(* IEC 61131-3 sources: plc-st-coding-agent/progress/evidence/f14_v14_remaining_20261113/jobs/custom_minimax-m27 (part 3) *)

(* ---- public-hard-05.raw_candidate_01.st ---- *)
(* ENGINEERING_CONTRACT - Mechanical Arm Control
 * =============================================================================
 * Mode Selection: Caller ensures exactly one mode active; emergency stop has highest priority.
 *
 * Output State Table:
 * | Output          | Activation                              | Retention                     | Reset                        | Priority    |
 * |-----------------|-----------------------------------------|-------------------------------|--------------------------------|-------------|
 * | MoveDown        | Manual:DownButton AND NOT DownLimitSwitch| Manual:button hold; Auto:step | EmergencyStop, step change   | Physical dir |
 * |                 | Auto: current step = down step           | Auto: hold until limit        | button release (manual)       | rule applies |
 * | MoveUp          | Manual:UpButton AND NOT UpLimitSwitch    | Manual:button hold; Auto:step | EmergencyStop, step change   | Physical dir |
 * |                 | Auto: current step = up step             | Auto: hold until limit        | button release (manual)       | rule applies |
 * | MoveLeft        | Manual:LeftButton AND NOT LeftLimitSwitch| Manual:button hold; Auto:step | EmergencyStop, step change   | Physical dir |
 * |                 | Auto: current step = left step           | Auto: hold until limit        | button release (manual)       | rule applies |
 * | MoveRight       | Manual:RightButton AND NOT RightLimitSwitch| Manual:button hold; Auto:step| EmergencyStop, step change   | Physical dir |
 * |                 | Auto: current step = right step          | Auto: hold until limit        | button release (manual)       | rule applies |
 * | ActivateGrip    | Manual:GripButton AND NOT GripLimitSwitch| Manual:button hold; Auto:step | EmergencyStop, step change   | N/A         |
 * |                 | Auto: grip step, hold until GripLimitSwitch| Auto: hold until limit       | button release (manual)       |             |
 * | ActivateRelease | Manual:ReleaseButton AND NOT ReleaseLimitSwitch| Manual:button hold; Auto:step| EmergencyStop, step change  | N/A         |
 * |                 | Auto: release step, hold until ReleaseLimitSwitch| Auto: hold until limit    | button release (manual)       |             |
 *
 * Sequence (8 steps, single cycle and continuous modes):
 *   0: Down -> 1: Grip -> 2: Up -> 3: Right -> 4: Down -> 5: Release -> 6: Up -> 7: Left -> (repeat)
 *
 * Single step mode: Same 8-step sequence, advancing one step per Start rising edge.
 * Single cycle mode: Executes all 8 steps, stops at stepIndex=8.
 * Continuous mode: Executes all 8 steps, returns to stepIndex=0 when complete.
 *
 * Units: Limit switches TRUE=at position (normally-open, closed at position).
 * Boundary: stepIndex ∈ [0..8]; 8 = cycle complete state for single cycle mode.
 * Same-scan: Final output evaluated from current stepIndex and limit switches per scan.
 *
 * Contract PUB clauses: PUB001-PUB020 define all behavior above.
 *)

FUNCTION_BLOCK ArmController
VAR
    stepIndex : INT := 0;         // Current step in sequence (0-7), 8 = single cycle complete
    startButtonPrev : BOOL := FALSE; // Rising edge detection for Start button
    tmpRisingEdge : BOOL;
END_VAR

(* CONTRACT_RULES
[
  {"kind": "hold_until_reset", "output": "MoveDown", "set_input": "DownButton", "reset_input": null},
  {"kind": "hold_until_reset", "output": "MoveUp", "set_input": "UpButton", "reset_input": null},
  {"kind": "hold_until_reset", "output": "MoveLeft", "set_input": "LeftButton", "reset_input": null},
  {"kind": "hold_until_reset", "output": "MoveRight", "set_input": "RightButton", "reset_input": null},
  {"kind": "hold_until_reset", "output": "ActivateGrip", "set_input": "GripButton", "reset_input": null},
  {"kind": "hold_until_reset", "output": "ActivateRelease", "set_input": "ReleaseButton", "reset_input": null}
]
*)

    // Emergency stop has highest priority - stops all outputs
    IF EmergencyStop = FALSE THEN
        MoveDown := FALSE;
        MoveUp := FALSE;
        MoveLeft := FALSE;
        MoveRight := FALSE;
        ActivateGrip := FALSE;
        ActivateRelease := FALSE;
    ELSIF SingleStepMode THEN
        // Detect rising edge on Start button
        tmpRisingEdge := Start AND NOT startButtonPrev;
        startButtonPrev := Start;

        IF tmpRisingEdge THEN
            stepIndex := stepIndex + 1;
            IF stepIndex > 7 THEN
                stepIndex := 0;
            END_IF
        END_IF

        // Execute current step
        CASE stepIndex OF
            0: // Down
                MoveDown := TRUE;
                IF DownLimitSwitch THEN
                    stepIndex := 1;
                END_IF
            1: // Grip
                ActivateGrip := TRUE;
                IF GripLimitSwitch THEN
                    stepIndex := 2;
                END_IF
            2: // Up
                MoveUp := TRUE;
                IF UpLimitSwitch THEN
                    stepIndex := 3;
                END_IF
            3: // Right
                MoveRight := TRUE;
                IF RightLimitSwitch THEN
                    stepIndex := 4;
                END_IF
            4: // Down (second descent)
                MoveDown := TRUE;
                IF DownLimitSwitch THEN
                    stepIndex := 5;
                END_IF
            5: // Release
                ActivateRelease := TRUE;
                IF ReleaseLimitSwitch THEN
                    stepIndex := 6;
                END_IF
            6: // Up (second ascent)
                MoveUp := TRUE;
                IF UpLimitSwitch THEN
                    stepIndex := 7;
                END_IF
            7: // Left (return to start)
                MoveLeft := TRUE;
                IF LeftLimitSwitch THEN
                    stepIndex := 0;
                END_IF
        END_CASE

    ELSIF SingleCycleMode THEN
        // Single cycle mode: run through all steps automatically, stop at end
        CASE stepIndex OF
            0:
                MoveDown := NOT DownLimitSwitch;
                IF DownLimitSwitch THEN
                    stepIndex := 1;
                END_IF
            1:
                ActivateGrip := NOT GripLimitSwitch;
                IF GripLimitSwitch THEN
                    stepIndex := 2;
                END_IF
            2:
                MoveUp := NOT UpLimitSwitch;
                IF UpLimitSwitch THEN
                    stepIndex := 3;
                END_IF
            3:
                MoveRight := NOT RightLimitSwitch;
                IF RightLimitSwitch THEN
                    stepIndex := 4;
                END_IF
            4:
                MoveDown := NOT DownLimitSwitch;
                IF DownLimitSwitch THEN
                    stepIndex := 5;
                END_IF
            5:
                ActivateRelease := NOT ReleaseLimitSwitch;
                IF ReleaseLimitSwitch THEN
                    stepIndex := 6;
                END_IF
            6:
                MoveUp := NOT UpLimitSwitch;
                IF UpLimitSwitch THEN
                    stepIndex := 7;
                END_IF
            7:
                MoveLeft := NOT LeftLimitSwitch;
                IF LeftLimitSwitch THEN
                    stepIndex := 8; // Cycle complete, stay here
                END_IF
        END_CASE

    ELSIF ContinuousMode THEN
        // Continuous mode: run through all steps automatically, restart at end
        CASE stepIndex OF
            0:
                MoveDown := NOT DownLimitSwitch;
                IF DownLimitSwitch THEN
                    stepIndex := 1;
                END_IF
            1:
                ActivateGrip := NOT GripLimitSwitch;
                IF GripLimitSwitch THEN
                    stepIndex := 2;
                END_IF
            2:
                MoveUp := NOT UpLimitSwitch;
                IF UpLimitSwitch THEN
                    stepIndex := 3;
                END_IF
            3:
                MoveRight := NOT RightLimitSwitch;
                IF RightLimitSwitch THEN
                    stepIndex := 4;
                END_IF
            4:
                MoveDown := NOT DownLimitSwitch;
                IF DownLimitSwitch THEN
                    stepIndex := 5;
                END_IF
            5:
                ActivateRelease := NOT ReleaseLimitSwitch;
                IF ReleaseLimitSwitch THEN
                    stepIndex := 6;
                END_IF
            6:
                MoveUp := NOT UpLimitSwitch;
                IF UpLimitSwitch THEN
                    stepIndex := 7;
                END_IF
            7:
                MoveLeft := NOT LeftLimitSwitch;
                IF LeftLimitSwitch THEN
                    stepIndex := 0; // Restart cycle
                END_IF
        END_CASE

    ELSIF ManualMode THEN
        // Manual mode: direct button control with limit switch protection
        MoveDown := DownButton AND NOT DownLimitSwitch;
        MoveUp := UpButton AND NOT UpLimitSwitch;
        MoveLeft := LeftButton AND NOT LeftLimitSwitch;
        MoveRight := RightButton AND NOT RightLimitSwitch;
        ActivateGrip := GripButton AND NOT GripLimitSwitch;
        ActivateRelease := ReleaseButton AND NOT ReleaseLimitSwitch;
    END_IF

END_FUNCTION_BLOCK

(* ---- public-hard-05.raw_candidate_02.st ---- *)
(* ENGINEERING_CONTRACT - Mechanical Arm Control
 * =============================================================================
 * Mode Selection: Caller ensures exactly one mode active; emergency stop has highest priority.
 *
 * Output State Table:
 * | Output          | Activation                              | Retention                     | Reset                        | Priority    |
 * |-----------------|-----------------------------------------|-------------------------------|--------------------------------|-------------|
 * | MoveDown        | Manual:DownButton AND NOT DownLimitSwitch| Manual:button hold; Auto:step | EmergencyStop, step change   | Physical dir |
 * |                 | Auto: current step = down step           | Auto: hold until limit        | button release (manual)       | rule applies |
 * | MoveUp          | Manual:UpButton AND NOT UpLimitSwitch    | Manual:button hold; Auto:step | EmergencyStop, step change   | Physical dir |
 * |                 | Auto: current step = up step             | Auto: hold until limit        | button release (manual)       | rule applies |
 * | MoveLeft        | Manual:LeftButton AND NOT LeftLimitSwitch| Manual:button hold; Auto:step | EmergencyStop, step change   | Physical dir |
 * |                 | Auto: current step = left step           | Auto: hold until limit        | button release (manual)       | rule applies |
 * | MoveRight       | Manual:RightButton AND NOT RightLimitSwitch| Manual:button hold; Auto:step| EmergencyStop, step change   | Physical dir |
 * |                 | Auto: current step = right step          | Auto: hold until limit        | button release (manual)       | rule applies |
 * | ActivateGrip    | Manual:GripButton AND NOT GripLimitSwitch| Manual:button hold; Auto:step | EmergencyStop, step change   | N/A         |
 * |                 | Auto: grip step, hold until GripLimitSwitch| Auto: hold until limit       | button release (manual)       |             |
 * | ActivateRelease | Manual:ReleaseButton AND NOT ReleaseLimitSwitch| Manual:button hold; Auto:step| EmergencyStop, step change  | N/A         |
 * |                 | Auto: release step, hold until ReleaseLimitSwitch| Auto: hold until limit    | button release (manual)       |             |
 *
 * Sequence (8 steps, single cycle and continuous modes):
 *   0: Down -> 1: Grip -> 2: Up -> 3: Right -> 4: Down -> 5: Release -> 6: Up -> 7: Left -> (repeat)
 *
 * Single step mode: Same 8-step sequence, advancing one step per Start rising edge.
 * Single cycle mode: Executes all 8 steps, stops at stepIndex=8.
 * Continuous mode: Executes all 8 steps, returns to stepIndex=0 when complete.
 *
 * Units: Limit switches TRUE=at position (normally-open, closed at position).
 * Boundary: stepIndex ∈ [0..8]; 8 = cycle complete state for single cycle mode.
 * Same-scan: Final output evaluated from current stepIndex and limit switches per scan.
 *
 * Contract PUB clauses: PUB001-PUB020 define all behavior above.
 *)

FUNCTION_BLOCK ArmController
VAR_INPUT
    ManualMode : BOOL;
    SingleStepMode : BOOL;
    SingleCycleMode : BOOL;
    ContinuousMode : BOOL;
    EmergencyStop : BOOL;
    Start : BOOL;
    DownButton : BOOL;
    UpButton : BOOL;
    LeftButton : BOOL;
    RightButton : BOOL;
    GripButton : BOOL;
    ReleaseButton : BOOL;
    DownLimitSwitch : BOOL;
    UpLimitSwitch : BOOL;
    LeftLimitSwitch : BOOL;
    RightLimitSwitch : BOOL;
    GripLimitSwitch : BOOL;
    ReleaseLimitSwitch : BOOL;
END_VAR
VAR_OUTPUT
    MoveDown : BOOL;
    MoveUp : BOOL;
    MoveLeft : BOOL;
    MoveRight : BOOL;
    ActivateGrip : BOOL;
    ActivateRelease : BOOL;
END_VAR
VAR
    stepIndex : INT := 0;         // Current step in sequence (0-7), 8 = single cycle complete
    startButtonPrev : BOOL := FALSE; // Rising edge detection for Start button
    tmpRisingEdge : BOOL;
END_VAR

(* CONTRACT_RULES
[
  {"kind": "hold_until_reset", "output": "MoveDown", "set_input": "DownButton", "reset_input": null},
  {"kind": "hold_until_reset", "output": "MoveUp", "set_input": "UpButton", "reset_input": null},
  {"kind": "hold_until_reset", "output": "MoveLeft", "set_input": "LeftButton", "reset_input": null},
  {"kind": "hold_until_reset", "output": "MoveRight", "set_input": "RightButton", "reset_input": null},
  {"kind": "hold_until_reset", "output": "ActivateGrip", "set_input": "GripButton", "reset_input": null},
  {"kind": "hold_until_reset", "output": "ActivateRelease", "set_input": "ReleaseButton", "reset_input": null}
]
*)

    // Emergency stop has highest priority - stops all outputs
    IF EmergencyStop = FALSE THEN
        MoveDown := FALSE;
        MoveUp := FALSE;
        MoveLeft := FALSE;
        MoveRight := FALSE;
        ActivateGrip := FALSE;
        ActivateRelease := FALSE;
    ELSIF SingleStepMode THEN
        // Detect rising edge on Start button
        tmpRisingEdge := Start AND NOT startButtonPrev;
        startButtonPrev := Start;

        IF tmpRisingEdge THEN
            stepIndex := stepIndex + 1;
            IF stepIndex > 7 THEN
                stepIndex := 0;
            END_IF;
        END_IF;

        // Execute current step
        CASE stepIndex OF
            0: // Down
                MoveDown := TRUE;
                IF DownLimitSwitch THEN
                    stepIndex := 1;
                END_IF;
            1: // Grip
                ActivateGrip := TRUE;
                IF GripLimitSwitch THEN
                    stepIndex := 2;
                END_IF;
            2: // Up
                MoveUp := TRUE;
                IF UpLimitSwitch THEN
                    stepIndex := 3;
                END_IF;
            3: // Right
                MoveRight := TRUE;
                IF RightLimitSwitch THEN
                    stepIndex := 4;
                END_IF;
            4: // Down (second descent)
                MoveDown := TRUE;
                IF DownLimitSwitch THEN
                    stepIndex := 5;
                END_IF;
            5: // Release
                ActivateRelease := TRUE;
                IF ReleaseLimitSwitch THEN
                    stepIndex := 6;
                END_IF;
            6: // Up (second ascent)
                MoveUp := TRUE;
                IF UpLimitSwitch THEN
                    stepIndex := 7;
                END_IF;
            7: // Left (return to start)
                MoveLeft := TRUE;
                IF LeftLimitSwitch THEN
                    stepIndex := 0;
                END_IF;
        END_CASE;

    ELSIF SingleCycleMode THEN
        // Single cycle mode: run through all steps automatically, stop at end
        CASE stepIndex OF
            0:
                MoveDown := NOT DownLimitSwitch;
                IF DownLimitSwitch THEN
                    stepIndex := 1;
                END_IF;
            1:
                ActivateGrip := NOT GripLimitSwitch;
                IF GripLimitSwitch THEN
                    stepIndex := 2;
                END_IF;
            2:
                MoveUp := NOT UpLimitSwitch;
                IF UpLimitSwitch THEN
                    stepIndex := 3;
                END_IF;
            3:
                MoveRight := NOT RightLimitSwitch;
                IF RightLimitSwitch THEN
                    stepIndex := 4;
                END_IF;
            4:
                MoveDown := NOT DownLimitSwitch;
                IF DownLimitSwitch THEN
                    stepIndex := 5;
                END_IF;
            5:
                ActivateRelease := NOT ReleaseLimitSwitch;
                IF ReleaseLimitSwitch THEN
                    stepIndex := 6;
                END_IF;
            6:
                MoveUp := NOT UpLimitSwitch;
                IF UpLimitSwitch THEN
                    stepIndex := 7;
                END_IF;
            7:
                MoveLeft := NOT LeftLimitSwitch;
                IF LeftLimitSwitch THEN
                    stepIndex := 8; // Cycle complete, stay here
                END_IF;
        END_CASE;

    ELSIF ContinuousMode THEN
        // Continuous mode: run through all steps automatically, restart at end
        CASE stepIndex OF
            0:
                MoveDown := NOT DownLimitSwitch;
                IF DownLimitSwitch THEN
                    stepIndex := 1;
                END_IF;
            1:
                ActivateGrip := NOT GripLimitSwitch;
                IF GripLimitSwitch THEN
                    stepIndex := 2;
                END_IF;
            2:
                MoveUp := NOT UpLimitSwitch;
                IF UpLimitSwitch THEN
                    stepIndex := 3;
                END_IF;
            3:
                MoveRight := NOT RightLimitSwitch;
                IF RightLimitSwitch THEN
                    stepIndex := 4;
                END_IF;
            4:
                MoveDown := NOT DownLimitSwitch;
                IF DownLimitSwitch THEN
                    stepIndex := 5;
                END_IF;
            5:
                ActivateRelease := NOT ReleaseLimitSwitch;
                IF ReleaseLimitSwitch THEN
                    stepIndex := 6;
                END_IF;
            6:
                MoveUp := NOT UpLimitSwitch;
                IF UpLimitSwitch THEN
                    stepIndex := 7;
                END_IF;
            7:
                MoveLeft := NOT LeftLimitSwitch;
                IF LeftLimitSwitch THEN
                    stepIndex := 0; // Restart cycle
                END_IF;
        END_CASE;

    ELSIF ManualMode THEN
        // Manual mode: direct button control with limit switch protection
        MoveDown := DownButton AND NOT DownLimitSwitch;
        MoveUp := UpButton AND NOT UpLimitSwitch;
        MoveLeft := LeftButton AND NOT LeftLimitSwitch;
        MoveRight := RightButton AND NOT RightLimitSwitch;
        ActivateGrip := GripButton AND NOT GripLimitSwitch;
        ActivateRelease := ReleaseButton AND NOT ReleaseLimitSwitch;
    END_IF;

END_FUNCTION_BLOCK

(* ---- public-hard-06.candidate_01.st ---- *)
FUNCTION_BLOCK ProductionControl
VAR_INPUT
    Mode            : BOOL;
    ForwardButton   : BOOL;
    ReverseButton   : BOOL;
    SensorFeed      : BOOL;
    SensorWash      : BOOL;
    SensorWeight    : BOOL;
    SensorFiring    : BOOL;
    SensorOutput    : BOOL;
    washComplete    : BOOL;
    weightComplete  : BOOL;
    weight          : REAL;
    firingComplete  : BOOL;
END_VAR
VAR_OUTPUT
    MotorForward    : BOOL;
    MotorReverse    : BOOL;
    kick             : BOOL;
    CompletionLight : BOOL;
    firingTemp      : REAL;
END_VAR
VAR
    eState          : INT := 0;
    tmp_WashTrig    : R_TRIG;
    tmp_WeightTrig  : R_TRIG;
    tmp_FiringTrig  : R_TRIG;
    tmp_FeedPrev    : BOOL := FALSE;
END_VAR

(*
ENGINEERING_CONTRACT
================================================================================
PUB001: Mode switch (0=manual, 1=automatic)
PUB002: Manual interlocks prevent simultaneous Forward/Reverse; priority=inhibit both
PUB003: Auto sequence: FEED→WASH→WEIGH→FIRING→OUTPUT→IDLE (reset on next SensorFeed)
PUB004: Weight check [100,200]; unqualified→kick=TRUE; qualified→firingTemp=(weight-100)*0.5+500
PUB006: washComplete starts MotorForward (rising-edge, state WASH)
PUB007: weightComplete triggers weight evaluation and either kick or motor start (rising-edge)
PUB008: firingComplete starts MotorForward (rising-edge, state FIRING)
PUB010: CompletionLight := SensorOutput (retention on product presence)
PUB012: Motor stops on sensor arrival; motor starts on completion signal or qualified weight
================================================================================
Output activation table:
| Output         | Set condition                              | Reset condition        |
|----------------|--------------------------------------------|------------------------|
| MotorForward   | SensorFeed in IDLE; washComplete in WASH;  | Sensor at next station;|
|                | weightComplete in WEIGH when qualified;    | Mode change;           |
|                | firingComplete in FIRING                   | IDLE;                  |
| MotorReverse   | ReverseButton AND NOT ForwardButton; Mode=0| Mode!=0; ForwardButton |
| kick           | weightComplete in WEIGH when unqualified   | Mode change; WEIGH entry|
| CompletionLight| SensorOutput=TRUE in OUTPUT                | SensorOutput=FALSE;Mode|
| firingTemp     | weightComplete in WEIGH when qualified     | Mode change; WEIGH entry|
================================================================================
*)

tmp_FeedPrev := SensorFeed;

CASE eState OF
    0: // IDLE
        MotorForward := FALSE;
        MotorReverse := FALSE;
        kick := FALSE;
        firingTemp := 0.0;
        IF Mode = FALSE THEN
            MotorForward := ForwardButton;
            MotorReverse := (NOT ForwardButton) AND ReverseButton;
        ELSE
            IF SensorFeed AND NOT tmp_FeedPrev THEN
                MotorForward := TRUE;
                eState := 1;
            END_IF;
        END_IF;

    1: // WASH
        IF Mode = FALSE THEN
            MotorForward := FALSE;
            MotorReverse := FALSE;
            kick := FALSE;
            firingTemp := 0.0;
            eState := 0;
        ELSE
            kick := FALSE;
            firingTemp := 0.0;
            tmp_WashTrig(CLK := washComplete);
            IF SensorWash THEN
                MotorForward := FALSE;
            END_IF;
            IF tmp_WashTrig.Q THEN
                MotorForward := TRUE;
                eState := 2;
            END_IF;
        END_IF;

    2: // WEIGH
        IF Mode = FALSE THEN
            MotorForward := FALSE;
            MotorReverse := FALSE;
            kick := FALSE;
            firingTemp := 0.0;
            eState := 0;
        ELSE
            IF SensorWeight THEN
                MotorForward := FALSE;
            END_IF;
            tmp_WeightTrig(CLK := weightComplete);
            IF tmp_WeightTrig.Q THEN
                IF (weight >= 100.0) AND (weight <= 200.0) THEN
                    firingTemp := (weight - 100.0) * 0.5 + 500.0;
                    kick := FALSE;
                    MotorForward := TRUE;
                    eState := 3;
                ELSE
                    kick := TRUE;
                    firingTemp := 0.0;
                    MotorForward := TRUE;
                    eState := 3;
                END_IF;
            END_IF;
        END_IF;

    3: // FIRING
        IF Mode = FALSE THEN
            MotorForward := FALSE;
            MotorReverse := FALSE;
            kick := FALSE;
            firingTemp := 0.0;
            eState := 0;
        ELSE
            IF SensorFiring THEN
                MotorForward := FALSE;
            END_IF;
            tmp_FiringTrig(CLK := firingComplete);
            IF tmp_FiringTrig.Q THEN
                MotorForward := TRUE;
                eState := 4;
            END_IF;
        END_IF;

    4: // OUTPUT
        IF Mode = FALSE THEN
            MotorForward := FALSE;
            MotorReverse := FALSE;
            kick := FALSE;
            firingTemp := 0.0;
            CompletionLight := FALSE;
            eState := 0;
        ELSE
            IF SensorOutput THEN
                MotorForward := FALSE;
                CompletionLight := TRUE;
            ELSE
                CompletionLight := FALSE;
            END_IF;
            IF NOT SensorOutput AND (NOT MotorForward) THEN
                eState := 0;
            END_IF;
        END_IF;
END_CASE;

(* CONTRACT_RULES
[
  {"kind": "hold_until_reset", "output": "kick", "set_input": "weightComplete", "reset_input": null},
  {"kind": "hold_until_reset", "output": "firingTemp", "set_input": "weightComplete", "reset_input": null}
]
*)
END_FUNCTION_BLOCK

(* ---- public-hard-06.patch_base_02.st ---- *)
FUNCTION_BLOCK ProductionControl
VAR_INPUT
    Mode            : BOOL;
    ForwardButton   : BOOL;
    ReverseButton   : BOOL;
    SensorFeed      : BOOL;
    SensorWash      : BOOL;
    SensorWeight    : BOOL;
    SensorFiring    : BOOL;
    SensorOutput    : BOOL;
    washComplete    : BOOL;
    weightComplete  : BOOL;
    weight          : REAL;
    firingComplete  : BOOL;
END_VAR
VAR_OUTPUT
    MotorForward    : BOOL;
    MotorReverse    : BOOL;
    kick             : BOOL;
    CompletionLight : BOOL;
    firingTemp      : REAL;
END_VAR
VAR
    eState          : INT := 0;
    tmp_WashTrig    : R_TRIG;
    tmp_WeightTrig  : R_TRIG;
    tmp_FiringTrig  : R_TRIG;
    tmp_FeedPrev    : BOOL := FALSE;
END_VAR

(*
ENGINEERING_CONTRACT
================================================================================
PUB001: Mode switch (0=manual, 1=automatic)
PUB002: Manual interlocks prevent simultaneous Forward/Reverse; priority=inhibit both
PUB003: Auto sequence: FEED→WASH→WEIGH→FIRING→OUTPUT→IDLE (reset on next SensorFeed)
PUB004: Weight check [100,200]; unqualified→kick=TRUE; qualified→firingTemp=(weight-100)*0.5+500
PUB006: washComplete starts MotorForward (rising-edge, state WASH)
PUB007: weightComplete triggers weight evaluation and either kick or motor start (rising-edge)
PUB008: firingComplete starts MotorForward (rising-edge, state FIRING)
PUB010: CompletionLight := SensorOutput (retention on product presence)
PUB012: Motor stops on sensor arrival; motor starts on completion signal or qualified weight
================================================================================
Output activation table:
| Output         | Set condition                              | Reset condition        |
|----------------|--------------------------------------------|------------------------|
| MotorForward   | SensorFeed in IDLE; washComplete in WASH;  | Sensor at next station;|
|                | weightComplete in WEIGH when qualified;    | Mode change;           |
|                | firingComplete in FIRING                   | IDLE;                  |
| MotorReverse   | ReverseButton AND NOT ForwardButton; Mode=0| Mode!=0; ForwardButton |
| kick           | weightComplete in WEIGH when unqualified   | Mode change; WEIGH entry|
| CompletionLight| SensorOutput=TRUE in OUTPUT                | SensorOutput=FALSE;Mode|
| firingTemp     | weightComplete in WEIGH when qualified     | Mode change; WEIGH entry|
================================================================================
*)

tmp_FeedPrev := SensorFeed;

CASE eState OF
    0: // IDLE
        MotorForward := FALSE;
        MotorReverse := FALSE;
        kick := FALSE;
        firingTemp := 0.0;
        IF Mode = FALSE THEN
            MotorForward := ForwardButton;
            MotorReverse := (NOT ForwardButton) AND ReverseButton;
        ELSE
            IF SensorFeed AND NOT tmp_FeedPrev THEN
                MotorForward := TRUE;
                eState := 1;
            END_IF;
        END_IF;

    1: // WASH
        IF Mode = FALSE THEN
            MotorForward := FALSE;
            MotorReverse := FALSE;
            kick := FALSE;
            firingTemp := 0.0;
            eState := 0;
        ELSE
            kick := FALSE;
            firingTemp := 0.0;
            tmp_WashTrig(CLK := washComplete);
            IF SensorWash THEN
                MotorForward := FALSE;
            END_IF;
            IF tmp_WashTrig.Q THEN
                MotorForward := TRUE;
                eState := 2;
            END_IF;
        END_IF;

    2: // WEIGH
        IF Mode = FALSE THEN
            MotorForward := FALSE;
            MotorReverse := FALSE;
            kick := FALSE;
            firingTemp := 0.0;
            eState := 0;
        ELSE
            IF SensorWeight THEN
                MotorForward := FALSE;
            END_IF;
            tmp_WeightTrig(CLK := weightComplete);
            IF tmp_WeightTrig.Q THEN
                IF (weight >= 100.0) AND (weight <= 200.0) THEN
                    firingTemp := (weight - 100.0) * 0.5 + 500.0;
                    kick := FALSE;
                    MotorForward := TRUE;
                    eState := 3;
                ELSE
                    kick := TRUE;
                    firingTemp := 0.0;
                    MotorForward := TRUE;
                    eState := 3;
                END_IF;
            END_IF;
        END_IF;

    3: // FIRING
        IF Mode = FALSE THEN
            MotorForward := FALSE;
            MotorReverse := FALSE;
            kick := FALSE;
            firingTemp := 0.0;
            eState := 0;
        ELSE
            IF SensorFiring THEN
                MotorForward := FALSE;
            END_IF;
            tmp_FiringTrig(CLK := firingComplete);
            IF tmp_FiringTrig.Q THEN
                MotorForward := TRUE;
                eState := 4;
            END_IF;
        END_IF;

    4: // OUTPUT
        IF Mode = FALSE THEN
            MotorForward := FALSE;
            MotorReverse := FALSE;
            kick := FALSE;
            firingTemp := 0.0;
            CompletionLight := FALSE;
            eState := 0;
        ELSE
            IF SensorOutput THEN
                MotorForward := FALSE;
                CompletionLight := TRUE;
            ELSE
                CompletionLight := FALSE;
            END_IF;
            IF NOT SensorOutput AND (NOT MotorForward) THEN
                eState := 0;
            END_IF;
        END_IF;
END_CASE;

(* CONTRACT_RULES
[
  {"kind": "hold_until_reset", "output": "kick", "set_input": "weightComplete", "reset_input": null},
  {"kind": "hold_until_reset", "output": "firingTemp", "set_input": "weightComplete", "reset_input": null}
]
*)
END_FUNCTION_BLOCK

(* ---- public-hard-06.patch_base_03.st ---- *)
FUNCTION_BLOCK ProductionControl
VAR_INPUT
    Mode            : BOOL;
    ForwardButton   : BOOL;
    ReverseButton   : BOOL;
    SensorFeed      : BOOL;
    SensorWash      : BOOL;
    SensorWeight    : BOOL;
    SensorFiring    : BOOL;
    SensorOutput    : BOOL;
    washComplete    : BOOL;
    weightComplete  : BOOL;
    weight          : REAL;
    firingComplete  : BOOL;
END_VAR
VAR_OUTPUT
    MotorForward    : BOOL;
    MotorReverse    : BOOL;
    kick             : BOOL;
    CompletionLight : BOOL;
    firingTemp      : REAL;
END_VAR
VAR
    eState          : INT := 0;
    tmp_WashTrig    : R_TRIG;
    tmp_WeightTrig  : R_TRIG;
    tmp_FiringTrig  : R_TRIG;
    tmp_FeedPrev    : BOOL := FALSE;
END_VAR

(*
ENGINEERING_CONTRACT
================================================================================
PUB001: Mode switch (0=manual, 1=automatic)
PUB002: Manual interlocks prevent simultaneous Forward/Reverse; priority=inhibit both
PUB003: Auto sequence: FEED→WASH→WEIGH→FIRING→OUTPUT→IDLE (reset on next SensorFeed)
PUB004: Weight check [100,200]; unqualified→kick=TRUE; qualified→firingTemp=(weight-100)*0.5+500
PUB006: washComplete starts MotorForward (rising-edge, state WASH)
PUB007: weightComplete triggers weight evaluation and either kick or motor start (rising-edge)
PUB008: firingComplete starts MotorForward (rising-edge, state FIRING)
PUB010: CompletionLight := SensorOutput (retention on product presence)
PUB012: Motor stops on sensor arrival; motor starts on completion signal or qualified weight
================================================================================
Output activation table:
| Output         | Set condition                              | Reset condition        |
|----------------|--------------------------------------------|------------------------|
| MotorForward   | SensorFeed in IDLE; washComplete in WASH;  | Sensor at next station;|
|                | weightComplete in WEIGH when qualified;    | Mode change;           |
|                | firingComplete in FIRING                   | IDLE;                  |
| MotorReverse   | ReverseButton AND NOT ForwardButton; Mode=0| Mode!=0; ForwardButton |
| kick           | weightComplete in WEIGH when unqualified   | Mode change; WEIGH entry|
| CompletionLight| SensorOutput=TRUE in OUTPUT                | SensorOutput=FALSE;Mode|
| firingTemp     | weightComplete in WEIGH when qualified     | Mode change; WEIGH entry|
================================================================================
*)

tmp_FeedPrev := SensorFeed;

CASE eState OF
    0: // IDLE
        MotorForward := FALSE;
        MotorReverse := FALSE;
        kick := FALSE;
        firingTemp := 0.0;
        IF Mode = FALSE THEN
            MotorForward := ForwardButton;
            MotorReverse := (NOT ForwardButton) AND ReverseButton;
        ELSE
            IF SensorFeed AND NOT tmp_FeedPrev THEN
                MotorForward := TRUE;
                eState := 1;
            END_IF;
        END_IF;

    1: // WASH
        IF Mode = FALSE THEN
            MotorForward := FALSE;
            MotorReverse := FALSE;
            kick := FALSE;
            firingTemp := 0.0;
            eState := 0;
        ELSE
            kick := FALSE;
            firingTemp := 0.0;
            tmp_WashTrig(CLK := washComplete);
            IF SensorWash THEN
                MotorForward := FALSE;
            END_IF;
            IF tmp_WashTrig.Q THEN
                MotorForward := TRUE;
                eState := 2;
            END_IF;
        END_IF;

    2: // WEIGH
        IF Mode = FALSE THEN
            MotorForward := FALSE;
            MotorReverse := FALSE;
            kick := FALSE;
            firingTemp := 0.0;
            eState := 0;
        ELSE
            IF SensorWeight THEN
                MotorForward := FALSE;
            END_IF;
            tmp_WeightTrig(CLK := weightComplete);
            IF tmp_WeightTrig.Q THEN
                IF (weight >= 100.0) AND (weight <= 200.0) THEN
                    firingTemp := (weight - 100.0) * 0.5 + 500.0;
                    kick := FALSE;
                    MotorForward := TRUE;
                    eState := 3;
                ELSE
                    kick := TRUE;
                    firingTemp := 0.0;
                    MotorForward := TRUE;
                    eState := 3;
                END_IF;
            END_IF;
        END_IF;

    3: // FIRING
        IF Mode = FALSE THEN
            MotorForward := FALSE;
            MotorReverse := FALSE;
            kick := FALSE;
            firingTemp := 0.0;
            eState := 0;
        ELSE
            IF SensorFiring THEN
                MotorForward := FALSE;
            END_IF;
            tmp_FiringTrig(CLK := firingComplete);
            IF tmp_FiringTrig.Q THEN
                MotorForward := TRUE;
                eState := 4;
            END_IF;
        END_IF;

    4: // OUTPUT
        IF Mode = FALSE THEN
            MotorForward := FALSE;
            MotorReverse := FALSE;
            kick := FALSE;
            firingTemp := 0.0;
            CompletionLight := FALSE;
            eState := 0;
        ELSE
            IF SensorOutput THEN
                MotorForward := FALSE;
                CompletionLight := TRUE;
            ELSE
                CompletionLight := FALSE;
            END_IF;
            IF NOT SensorOutput AND (NOT MotorForward) THEN
                eState := 0;
            END_IF;
        END_IF;
END_CASE;

(* CONTRACT_RULES
[
  {"kind": "hold_until_reset", "output": "kick", "set_input": "weightComplete", "reset_input": null},
  {"kind": "hold_until_reset", "output": "firingTemp", "set_input": "weightComplete", "reset_input": null}
]
*)
END_FUNCTION_BLOCK

(* ---- public-hard-06.raw_candidate_01.st ---- *)
FUNCTION_BLOCK ProductionControl
VAR_INPUT
    Mode            : BOOL;
    ForwardButton   : BOOL;
    ReverseButton   : BOOL;
    SensorFeed      : BOOL;
    SensorWash      : BOOL;
    SensorWeight    : BOOL;
    SensorFiring    : BOOL;
    SensorOutput    : BOOL;
    washComplete    : BOOL;
    weightComplete  : BOOL;
    weight          : REAL;
    firingComplete  : BOOL;
END_VAR
VAR_OUTPUT
    MotorForward    : BOOL;
    MotorReverse    : BOOL;
    kick             : BOOL;
    CompletionLight : BOOL;
    firingTemp      : REAL;
END_VAR
VAR
    eState          : INT := 0;
    tmp_WashTrig    : R_TRIG;
    tmp_WeightTrig  : R_TRIG;
    tmp_FiringTrig  : R_TRIG;
    tmp_FeedPrev    : BOOL := FALSE;
END_VAR

(*
ENGINEERING_CONTRACT
================================================================================
PUB001: Mode switch (0=manual, 1=automatic)
PUB002: Manual interlocks prevent simultaneous Forward/Reverse; priority=inhibit both
PUB003: Auto sequence: FEED→WASH→WEIGH→FIRING→OUTPUT→IDLE (reset on next SensorFeed)
PUB004: Weight check [100,200]; unqualified→kick=TRUE; qualified→firingTemp=(weight-100)*0.5+500
PUB006: washComplete starts MotorForward (rising-edge, state WASH)
PUB007: weightComplete triggers weight evaluation and either kick or motor start (rising-edge)
PUB008: firingComplete starts MotorForward (rising-edge, state FIRING)
PUB010: CompletionLight := SensorOutput (retention on product presence)
PUB012: Motor stops on sensor arrival; motor starts on completion signal or qualified weight
================================================================================
Output activation table:
| Output         | Set condition                              | Reset condition        |
|----------------|--------------------------------------------|------------------------|
| MotorForward   | SensorFeed in IDLE; washComplete in WASH;  | Sensor at next station;|
|                | weightComplete in WEIGH when qualified;    | Mode change;           |
|                | firingComplete in FIRING                   | IDLE;                  |
| MotorReverse   | ReverseButton AND NOT ForwardButton; Mode=0| Mode!=0; ForwardButton |
| kick           | weightComplete in WEIGH when unqualified   | Mode change; WEIGH entry|
| CompletionLight| SensorOutput=TRUE in OUTPUT                | SensorOutput=FALSE;Mode|
| firingTemp     | weightComplete in WEIGH when qualified     | Mode change; WEIGH entry|
================================================================================
*)

tmp_FeedPrev := SensorFeed;

CASE eState OF
    0: // IDLE
        MotorForward := FALSE;
        MotorReverse := FALSE;
        kick := FALSE;
        firingTemp := 0.0;
        IF Mode = FALSE THEN
            MotorForward := ForwardButton;
            MotorReverse := (NOT ForwardButton) AND ReverseButton;
        ELSE
            IF SensorFeed AND NOT tmp_FeedPrev THEN
                MotorForward := TRUE;
                eState := 1;
            END_IF;
        END_IF;

    1: // WASH
        IF Mode = FALSE THEN
            MotorForward := FALSE;
            MotorReverse := FALSE;
            kick := FALSE;
            firingTemp := 0.0;
            eState := 0;
        ELSE
            kick := FALSE;
            firingTemp := 0.0;
            tmp_WashTrig(CLK := washComplete);
            IF SensorWash THEN
                MotorForward := FALSE;
            END_IF;
            IF tmp_WashTrig.Q THEN
                MotorForward := TRUE;
                eState := 2;
            END_IF;
        END_IF;

    2: // WEIGH
        IF Mode = FALSE THEN
            MotorForward := FALSE;
            MotorReverse := FALSE;
            kick := FALSE;
            firingTemp := 0.0;
            eState := 0;
        ELSE
            IF SensorWeight THEN
                MotorForward := FALSE;
            END_IF;
            tmp_WeightTrig(CLK := weightComplete);
            IF tmp_WeightTrig.Q THEN
                IF (weight >= 100.0) AND (weight <= 200.0) THEN
                    firingTemp := (weight - 100.0) * 0.5 + 500.0;
                    kick := FALSE;
                    MotorForward := TRUE;
                    eState := 3;
                ELSE
                    kick := TRUE;
                    firingTemp := 0.0;
                    MotorForward := TRUE;
                    eState := 3;
                END_IF;
            END_IF;
        END_IF;

    3: // FIRING
        IF Mode = FALSE THEN
            MotorForward := FALSE;
            MotorReverse := FALSE;
            kick := FALSE;
            firingTemp := 0.0;
            eState := 0;
        ELSE
            IF SensorFiring THEN
                MotorForward := FALSE;
            END_IF;
            tmp_FiringTrig(CLK := firingComplete);
            IF tmp_FiringTrig.Q THEN
                MotorForward := TRUE;
                eState := 4;
            END_IF;
        END_IF;

    4: // OUTPUT
        IF Mode = FALSE THEN
            MotorForward := FALSE;
            MotorReverse := FALSE;
            kick := FALSE;
            firingTemp := 0.0;
            CompletionLight := FALSE;
            eState := 0;
        ELSE
            IF SensorOutput THEN
                MotorForward := FALSE;
                CompletionLight := TRUE;
            ELSE
                CompletionLight := FALSE;
            END_IF;
            IF NOT SensorOutput AND (NOT MotorForward) THEN
                eState := 0;
            END_IF;
        END_IF;
END_CASE;

(* CONTRACT_RULES
[
  {"kind": "hold_until_reset", "output": "kick", "set_input": "weightComplete", "reset_input": null},
  {"kind": "hold_until_reset", "output": "firingTemp", "set_input": "weightComplete", "reset_input": null}
]
*)
END_FUNCTION_BLOCK

(* ---- public-medium-01.candidate_01.st ---- *)
FUNCTION_BLOCK FB_PumpControl
VAR_INPUT
    mode  : BOOL;  // FALSE: Manual, TRUE: Automatic
    start : BOOL;
    stop  : BOOL;
END_VAR

VAR_IN_OUT
    pumpGroup : ARRAY[1..5] OF ST_Pump;
END_VAR

VAR
    tmp_i          : INT;
    tmp_j          : INT;
    tmp_temp       : ST_Pump;
    tmp_tempIndex  : INT;
    tmp_sorted     : ARRAY[1..5] OF ST_Pump;
    tmp_order      : ARRAY[1..5] OF INT;
END_VAR

// ENGINEERING_CONTRACT
// ┌─────────────────────────────────────────────────────────────────────────────────────────────┐
// │ Output/State              │ Activation                   │ Retention    │ Reset/Deactivation │ Same-scan │ Boundaries      │ PUB Clause     │
// │------------------------───│──────────────────────────────│──────────────│────────────────────│───────────│─────────────────│────────────────│
// │ pumpGroup[].RunComd FALSE │ stop=TRUE                    │ -            │ start=TRUE         │ -         │ 0–5 pumps       │ PUB001, PUB004 │
// │ pumpGroup[].RunComd TRUE  │ start=TRUE AND selected only │ Hold(start)  │ stop=TRUE          │ -         │ Manual: 1–5 pumps; Auto: 3 │ PUB001, PUB003 │
// │ pumpGroup[].RunComd TRUE  │ start=TRUE AND top-3 priority│ Hold(start)  │ stop=TRUE          │ -         │ Auto: exactly 3 │ PUB002         │
// └─────────────────────────────────────────────────────────────────────────────────────────────┘

// Stop has highest priority — de-energizes all pumps immediately
IF stop THEN
    FOR tmp_i := 1 TO 5 DO
        pumpGroup[tmp_i].RunComd := FALSE;
    END_FOR;
    RETURN;
END_IF;

IF NOT mode THEN
    // Manual mode: selected pump(s) follow start command
    FOR tmp_i := 1 TO 5 DO
        IF pumpGroup[tmp_i].selection THEN
            pumpGroup[tmp_i].RunComd := start;
        ELSE
            pumpGroup[tmp_i].RunComd := FALSE;
        END_IF;
    END_FOR;
ELSE
    // Automatic mode: top-3 priority pumps follow start command
    // Copy for sorting (preserves original pumpGroup indices)
    FOR tmp_i := 1 TO 5 DO
        tmp_sorted[tmp_i] := pumpGroup[tmp_i];
        tmp_order[tmp_i]  := tmp_i;
    END_FOR;

    // Bubble sort by priority descending (stable: equal priority keeps original order)
    FOR tmp_i := 1 TO 4 DO
        FOR tmp_j := tmp_i + 1 TO 5 DO
            IF tmp_sorted[tmp_j].priority > tmp_sorted[tmp_i].priority THEN
                tmp_temp           := tmp_sorted[tmp_i];
                tmp_sorted[tmp_i]  := tmp_sorted[tmp_j];
                tmp_sorted[tmp_j]  := tmp_temp;

                tmp_tempIndex      := tmp_order[tmp_i];
                tmp_order[tmp_i]   := tmp_order[tmp_j];
                tmp_order[tmp_j]   := tmp_tempIndex;
            END_IF;
        END_FOR;
    END_FOR;

    // Enable top-3 pumps (by original index) when start is asserted
    FOR tmp_i := 1 TO 5 DO
        IF tmp_i <= 3 THEN
            pumpGroup[tmp_order[tmp_i]].RunComd := start;
        ELSE
            pumpGroup[tmp_order[tmp_i]].RunComd := FALSE;
        END_IF;
    END_FOR;
END_IF;

END_FUNCTION_BLOCK

(* CONTRACT_RULES [] *)

(* ---- public-medium-01.candidate_02.st ---- *)
TYPE ST_Pump : STRUCT
    priority  : INT;
    selection : BOOL;
    RunComd   : BOOL;
END_STRUCT
END_TYPE;

FUNCTION_BLOCK FB_PumpControl
VAR_INPUT
    mode  : BOOL;  // FALSE: Manual, TRUE: Automatic
    start : BOOL;
    stop  : BOOL;
END_VAR

VAR_IN_OUT
    pumpGroup : ARRAY[1..5] OF ST_Pump;
END_VAR

VAR
    tmp_i          : INT;
    tmp_j          : INT;
    tmp_temp       : ST_Pump;
    tmp_tempIndex  : INT;
    tmp_sorted     : ARRAY[1..5] OF ST_Pump;
    tmp_order      : ARRAY[1..5] OF INT;
END_VAR

// ENGINEERING_CONTRACT
// ┌─────────────────────────────────────────────────────────────────────────────────────────────┐
// │ Output/State              │ Activation                   │ Retention    │ Reset/Deactivation │ Same-scan │ Boundaries      │ PUB Clause     │
// │------------------------───│──────────────────────────────│──────────────│────────────────────│───────────│─────────────────│────────────────│
// │ pumpGroup[].RunComd FALSE │ stop=TRUE                    │ -            │ start=TRUE         │ -         │ 0–5 pumps       │ PUB001, PUB004 │
// │ pumpGroup[].RunComd TRUE  │ start=TRUE AND selected only │ Hold(start)  │ stop=TRUE          │ -         │ Manual: 1–5 pumps; Auto: 3 │ PUB001, PUB003 │
// │ pumpGroup[].RunComd TRUE  │ start=TRUE AND top-3 priority│ Hold(start)  │ stop=TRUE          │ -         │ Auto: exactly 3 │ PUB002         │
// └─────────────────────────────────────────────────────────────────────────────────────────────┘

// Stop has highest priority — de-energizes all pumps immediately
IF stop THEN
    FOR tmp_i := 1 TO 5 DO
        pumpGroup[tmp_i].RunComd := FALSE;
    END_FOR;
    RETURN;
END_IF;

IF NOT mode THEN
    // Manual mode: selected pump(s) follow start command
    FOR tmp_i := 1 TO 5 DO
        IF pumpGroup[tmp_i].selection THEN
            pumpGroup[tmp_i].RunComd := start;
        ELSE
            pumpGroup[tmp_i].RunComd := FALSE;
        END_IF;
    END_FOR;
ELSE
    // Automatic mode: top-3 priority pumps follow start command
    // Copy for sorting (preserves original pumpGroup indices)
    FOR tmp_i := 1 TO 5 DO
        tmp_sorted[tmp_i] := pumpGroup[tmp_i];
        tmp_order[tmp_i]  := tmp_i;
    END_FOR;

    // Bubble sort by priority descending (stable: equal priority keeps original order)
    FOR tmp_i := 1 TO 4 DO
        FOR tmp_j := tmp_i + 1 TO 5 DO
            IF tmp_sorted[tmp_j].priority > tmp_sorted[tmp_i].priority THEN
                tmp_temp           := tmp_sorted[tmp_i];
                tmp_sorted[tmp_i]  := tmp_sorted[tmp_j];
                tmp_sorted[tmp_j]  := tmp_temp;

                tmp_tempIndex      := tmp_order[tmp_i];
                tmp_order[tmp_i]   := tmp_order[tmp_j];
                tmp_order[tmp_j]   := tmp_tempIndex;
            END_IF;
        END_FOR;
    END_FOR;

    // Enable top-3 pumps (by original index) when start is asserted
    FOR tmp_i := 1 TO 5 DO
        IF tmp_i <= 3 THEN
            pumpGroup[tmp_order[tmp_i]].RunComd := start;
        ELSE
            pumpGroup[tmp_order[tmp_i]].RunComd := FALSE;
        END_IF;
    END_FOR;
END_IF;

END_FUNCTION_BLOCK

(* CONTRACT_RULES [] *)

(* ---- public-medium-01.patch_base_02.st ---- *)
FUNCTION_BLOCK FB_PumpControl
VAR_INPUT
    mode  : BOOL;  // FALSE: Manual, TRUE: Automatic
    start : BOOL;
    stop  : BOOL;
END_VAR

VAR_IN_OUT
    pumpGroup : ARRAY[1..5] OF ST_Pump;
END_VAR

VAR
    tmp_i          : INT;
    tmp_j          : INT;
    tmp_temp       : ST_Pump;
    tmp_tempIndex  : INT;
    tmp_sorted     : ARRAY[1..5] OF ST_Pump;
    tmp_order      : ARRAY[1..5] OF INT;
END_VAR

// ENGINEERING_CONTRACT
// ┌─────────────────────────────────────────────────────────────────────────────────────────────┐
// │ Output/State              │ Activation                   │ Retention    │ Reset/Deactivation │ Same-scan │ Boundaries      │ PUB Clause     │
// │------------------------───│──────────────────────────────│──────────────│────────────────────│───────────│─────────────────│────────────────│
// │ pumpGroup[].RunComd FALSE │ stop=TRUE                    │ -            │ start=TRUE         │ -         │ 0–5 pumps       │ PUB001, PUB004 │
// │ pumpGroup[].RunComd TRUE  │ start=TRUE AND selected only │ Hold(start)  │ stop=TRUE          │ -         │ Manual: 1–5 pumps; Auto: 3 │ PUB001, PUB003 │
// │ pumpGroup[].RunComd TRUE  │ start=TRUE AND top-3 priority│ Hold(start)  │ stop=TRUE          │ -         │ Auto: exactly 3 │ PUB002         │
// └─────────────────────────────────────────────────────────────────────────────────────────────┘

// Stop has highest priority — de-energizes all pumps immediately
IF stop THEN
    FOR tmp_i := 1 TO 5 DO
        pumpGroup[tmp_i].RunComd := FALSE;
    END_FOR;
    RETURN;
END_IF;

IF NOT mode THEN
    // Manual mode: selected pump(s) follow start command
    FOR tmp_i := 1 TO 5 DO
        IF pumpGroup[tmp_i].selection THEN
            pumpGroup[tmp_i].RunComd := start;
        ELSE
            pumpGroup[tmp_i].RunComd := FALSE;
        END_IF;
    END_FOR;
ELSE
    // Automatic mode: top-3 priority pumps follow start command
    // Copy for sorting (preserves original pumpGroup indices)
    FOR tmp_i := 1 TO 5 DO
        tmp_sorted[tmp_i] := pumpGroup[tmp_i];
        tmp_order[tmp_i]  := tmp_i;
    END_FOR;

    // Bubble sort by priority descending (stable: equal priority keeps original order)
    FOR tmp_i := 1 TO 4 DO
        FOR tmp_j := tmp_i + 1 TO 5 DO
            IF tmp_sorted[tmp_j].priority > tmp_sorted[tmp_i].priority THEN
                tmp_temp           := tmp_sorted[tmp_i];
                tmp_sorted[tmp_i]  := tmp_sorted[tmp_j];
                tmp_sorted[tmp_j]  := tmp_temp;

                tmp_tempIndex      := tmp_order[tmp_i];
                tmp_order[tmp_i]   := tmp_order[tmp_j];
                tmp_order[tmp_j]   := tmp_tempIndex;
            END_IF;
        END_FOR;
    END_FOR;

    // Enable top-3 pumps (by original index) when start is asserted
    FOR tmp_i := 1 TO 5 DO
        IF tmp_i <= 3 THEN
            pumpGroup[tmp_order[tmp_i]].RunComd := start;
        ELSE
            pumpGroup[tmp_order[tmp_i]].RunComd := FALSE;
        END_IF;
    END_FOR;
END_IF;

END_FUNCTION_BLOCK

(* CONTRACT_RULES [] *)

(* ---- public-medium-01.raw_candidate_01.st ---- *)
FUNCTION_BLOCK FB_PumpControl
VAR_INPUT
    mode  : BOOL;  // FALSE: Manual, TRUE: Automatic
    start : BOOL;
    stop  : BOOL;
END_VAR

VAR_IN_OUT
    pumpGroup : ARRAY[1..5] OF ST_Pump;
END_VAR

VAR
    tmp_i          : INT;
    tmp_j          : INT;
    tmp_temp       : ST_Pump;
    tmp_tempIndex  : INT;
    tmp_sorted     : ARRAY[1..5] OF ST_Pump;
    tmp_order      : ARRAY[1..5] OF INT;
END_VAR

// ENGINEERING_CONTRACT
// ┌─────────────────────────────────────────────────────────────────────────────────────────────┐
// │ Output/State              │ Activation                   │ Retention    │ Reset/Deactivation │ Same-scan │ Boundaries      │ PUB Clause     │
// │------------------------───│──────────────────────────────│──────────────│────────────────────│───────────│─────────────────│────────────────│
// │ pumpGroup[].RunComd FALSE │ stop=TRUE                    │ -            │ start=TRUE         │ -         │ 0–5 pumps       │ PUB001, PUB004 │
// │ pumpGroup[].RunComd TRUE  │ start=TRUE AND selected only │ Hold(start)  │ stop=TRUE          │ -         │ Manual: 1–5 pumps; Auto: 3 │ PUB001, PUB003 │
// │ pumpGroup[].RunComd TRUE  │ start=TRUE AND top-3 priority│ Hold(start)  │ stop=TRUE          │ -         │ Auto: exactly 3 │ PUB002         │
// └─────────────────────────────────────────────────────────────────────────────────────────────┘

// Stop has highest priority — de-energizes all pumps immediately
IF stop THEN
    FOR tmp_i := 1 TO 5 DO
        pumpGroup[tmp_i].RunComd := FALSE;
    END_FOR
    RETURN;
END_IF

IF NOT mode THEN
    // Manual mode: selected pump(s) follow start command
    FOR tmp_i := 1 TO 5 DO
        IF pumpGroup[tmp_i].selection THEN
            pumpGroup[tmp_i].RunComd := start;
        ELSE
            pumpGroup[tmp_i].RunComd := FALSE;
        END_IF
    END_FOR
ELSE
    // Automatic mode: top-3 priority pumps follow start command
    // Copy for sorting (preserves original pumpGroup indices)
    FOR tmp_i := 1 TO 5 DO
        tmp_sorted[tmp_i] := pumpGroup[tmp_i];
        tmp_order[tmp_i]  := tmp_i;
    END_FOR

    // Bubble sort by priority descending (stable: equal priority keeps original order)
    FOR tmp_i := 1 TO 4 DO
        FOR tmp_j := tmp_i + 1 TO 5 DO
            IF tmp_sorted[tmp_j].priority > tmp_sorted[tmp_i].priority THEN
                tmp_temp           := tmp_sorted[tmp_i];
                tmp_sorted[tmp_i]  := tmp_sorted[tmp_j];
                tmp_sorted[tmp_j]  := tmp_temp;

                tmp_tempIndex      := tmp_order[tmp_i];
                tmp_order[tmp_i]   := tmp_order[tmp_j];
                tmp_order[tmp_j]   := tmp_tempIndex;
            END_IF
        END_FOR
    END_FOR

    // Enable top-3 pumps (by original index) when start is asserted
    FOR tmp_i := 1 TO 5 DO
        IF tmp_i <= 3 THEN
            pumpGroup[tmp_order[tmp_i]].RunComd := start;
        ELSE
            pumpGroup[tmp_order[tmp_i]].RunComd := FALSE;
        END_IF
    END_FOR
END_IF

END_FUNCTION_BLOCK

(* CONTRACT_RULES [] *)

(* ---- public-medium-01.raw_candidate_02.st ---- *)
TYPE ST_Pump : STRUCT
    priority  : INT;
    selection : BOOL;
    RunComd   : BOOL;
END_STRUCT
END_TYPE

FUNCTION_BLOCK FB_PumpControl
VAR_INPUT
    mode  : BOOL;  // FALSE: Manual, TRUE: Automatic
    start : BOOL;
    stop  : BOOL;
END_VAR

VAR_IN_OUT
    pumpGroup : ARRAY[1..5] OF ST_Pump;
END_VAR

VAR
    tmp_i          : INT;
    tmp_j          : INT;
    tmp_temp       : ST_Pump;
    tmp_tempIndex  : INT;
    tmp_sorted     : ARRAY[1..5] OF ST_Pump;
    tmp_order      : ARRAY[1..5] OF INT;
END_VAR

// ENGINEERING_CONTRACT
// ┌─────────────────────────────────────────────────────────────────────────────────────────────┐
// │ Output/State              │ Activation                   │ Retention    │ Reset/Deactivation │ Same-scan │ Boundaries      │ PUB Clause     │
// │------------------------───│──────────────────────────────│──────────────│────────────────────│───────────│─────────────────│────────────────│
// │ pumpGroup[].RunComd FALSE │ stop=TRUE                    │ -            │ start=TRUE         │ -         │ 0–5 pumps       │ PUB001, PUB004 │
// │ pumpGroup[].RunComd TRUE  │ start=TRUE AND selected only │ Hold(start)  │ stop=TRUE          │ -         │ Manual: 1–5 pumps; Auto: 3 │ PUB001, PUB003 │
// │ pumpGroup[].RunComd TRUE  │ start=TRUE AND top-3 priority│ Hold(start)  │ stop=TRUE          │ -         │ Auto: exactly 3 │ PUB002         │
// └─────────────────────────────────────────────────────────────────────────────────────────────┘

// Stop has highest priority — de-energizes all pumps immediately
IF stop THEN
    FOR tmp_i := 1 TO 5 DO
        pumpGroup[tmp_i].RunComd := FALSE;
    END_FOR;
    RETURN;
END_IF;

IF NOT mode THEN
    // Manual mode: selected pump(s) follow start command
    FOR tmp_i := 1 TO 5 DO
        IF pumpGroup[tmp_i].selection THEN
            pumpGroup[tmp_i].RunComd := start;
        ELSE
            pumpGroup[tmp_i].RunComd := FALSE;
        END_IF;
    END_FOR;
ELSE
    // Automatic mode: top-3 priority pumps follow start command
    // Copy for sorting (preserves original pumpGroup indices)
    FOR tmp_i := 1 TO 5 DO
        tmp_sorted[tmp_i] := pumpGroup[tmp_i];
        tmp_order[tmp_i]  := tmp_i;
    END_FOR;

    // Bubble sort by priority descending (stable: equal priority keeps original order)
    FOR tmp_i := 1 TO 4 DO
        FOR tmp_j := tmp_i + 1 TO 5 DO
            IF tmp_sorted[tmp_j].priority > tmp_sorted[tmp_i].priority THEN
                tmp_temp           := tmp_sorted[tmp_i];
                tmp_sorted[tmp_i]  := tmp_sorted[tmp_j];
                tmp_sorted[tmp_j]  := tmp_temp;

                tmp_tempIndex      := tmp_order[tmp_i];
                tmp_order[tmp_i]   := tmp_order[tmp_j];
                tmp_order[tmp_j]   := tmp_tempIndex;
            END_IF;
        END_FOR;
    END_FOR;

    // Enable top-3 pumps (by original index) when start is asserted
    FOR tmp_i := 1 TO 5 DO
        IF tmp_i <= 3 THEN
            pumpGroup[tmp_order[tmp_i]].RunComd := start;
        ELSE
            pumpGroup[tmp_order[tmp_i]].RunComd := FALSE;
        END_IF;
    END_FOR;
END_IF;

END_FUNCTION_BLOCK

(* CONTRACT_RULES [] *)

(* ---- public-medium-02.candidate_01.st ---- *)
FUNCTION_BLOCK FB_AnalogBatchProcessing
VAR_INPUT
END_VAR
VAR_IN_OUT
    analogValues : ARRAY[*] OF INT;
    channels     : ARRAY[*] OF ST_AnalogChannel;
END_VAR
VAR_OUTPUT
END_VAR
VAR
END_VAR

(*
ENGINEERING_CONTRACT
================================================================================
PUB001: Process 'count' channels starting at each array's lower bound.
        Arrays passed by reference preserve caller-defined bounds.
        Read-only: analogValues elements are never modified.
PUB002: Per-channel conversion based on measuringMode field.
        - Mode 0: Linear scaling using hiLIM/loLIM and bipolar flag.
        - Mode 1: Standard temperature (raw / 10.0).
        - Mode 2: Climatic temperature (raw / 100.0).
        - Invalid mode: retVal=16#8001, outputValue unchanged.
PUB003: Mode 0 linear scaling maps raw 0..27648 (unipolar) or -27648..27648 (bipolar)
        to loLIM..hiLIM range. OutputValue = loLIM + (raw - rawMin) * (hiLIM - loLIM) / range.
PUB004: If hiLIM <= loLIM in mode 0, set retVal=16#8002 and skip conversion.
PUB005: Disabled channels (enable=FALSE) are skipped; retVal and outputValue unchanged.
PUB006: Per-channel retVal WORD status: 16#8001 (invalid mode), 16#8002 (bad range).
PUB007: Same-scan priority: enable→measuringMode→hiLIM/loLIM check→conversion.
PUB008: Temperature output = raw / divisor (10 or 100) as REAL.
--------------------------------------------------------------------------------
*)

VAR
    tmpIndex     : DINT;
    tmpRaw       : INT;
    tmpRawReal   : REAL;
    tmpRange     : REAL;
    tmpOffset    : REAL;
    tmpChannel   : ST_AnalogChannel;
    tmpLower     : DINT;
    tmpUpperAna  : DINT;
    tmpUpperCh   : DINT;
    tmpProcessed : BOOL;
END_VAR

(* CONTRACT_RULES [] *)

tmpLower    := LOWER_BOUND(analogValues, 1);
tmpUpperAna := UPPER_BOUND(analogValues, 1);
tmpUpperCh  := UPPER_BOUND(channels, 1);

FOR tmpIndex := 0 TO (count - 1) DO
    tmpProcessed := FALSE;

    (* Bounds check: skip if index exceeds either array *)
    IF (tmpLower + tmpIndex) > tmpUpperAna OR (tmpLower + tmpIndex) > tmpUpperCh THEN
        CONTINUE;
    END_IF;

    tmpChannel := channels[tmpLower + tmpIndex];

    (* Skip disabled channels; retain previous outputValue and retVal *)
    IF NOT tmpChannel.enable THEN
        CONTINUE;
    END_IF;

    (* Determine conversion based on measuringMode *)
    IF tmpChannel.measuringMode = 0 THEN
        (* Non-temperature linear scaling *)
        IF tmpChannel.hiLIM <= tmpChannel.loLIM THEN
            channels[tmpLower + tmpIndex].retVal := 16#8002;
        ELSE
            tmpRaw       := analogValues[tmpLower + tmpIndex];
            tmpRawReal   := TO_REAL(tmpRaw);
            tmpRange     := tmpChannel.hiLIM - tmpChannel.loLIM;

            IF tmpChannel.bipolar THEN
                (* Map -27648..27648 to loLIM..hiLIM *)
                tmpOffset    := TO_REAL(27648);
                channels[tmpLower + tmpIndex].outputValue := tmpChannel.loLIM +
                    (tmpRawReal + tmpOffset) * tmpRange / TO_REAL(55296);
            ELSE
                (* Map 0..27648 to loLIM..hiLIM *)
                channels[tmpLower + tmpIndex].outputValue := tmpChannel.loLIM +
                    tmpRawReal * tmpRange / TO_REAL(27648);
            END_IF;
            channels[tmpLower + tmpIndex].retVal := 0;
        END_IF;
        tmpProcessed := TRUE;
    ELSIF tmpChannel.measuringMode = 1 THEN
        (* Standard temperature: outputValue = raw / 10 *)
        tmpRaw := analogValues[tmpLower + tmpIndex];
        channels[tmpLower + tmpIndex].outputValue := TO_REAL(tmpRaw) / TO_REAL(10);
        channels[tmpLower + tmpIndex].retVal := 0;
        tmpProcessed := TRUE;
    ELSIF tmpChannel.measuringMode = 2 THEN
        (* Climatic temperature: outputValue = raw / 100 *)
        tmpRaw := analogValues[tmpLower + tmpIndex];
        channels[tmpLower + tmpIndex].outputValue := TO_REAL(tmpRaw) / TO_REAL(100);
        channels[tmpLower + tmpIndex].retVal := 0;
        tmpProcessed := TRUE;
    END_IF;

    (* Invalid measuringMode (not 0, 1, or 2) *)
    IF NOT tmpProcessed THEN
        channels[tmpLower + tmpIndex].retVal := 16#8001;
    END_IF;

END_FOR;

END_FUNCTION_BLOCK

(* ---- public-medium-02.candidate_02.st ---- *)
TYPE ST_AnalogChannel :
STRUCT
    enable         : BOOL;
    hiLIM          : REAL;
    loLIM          : REAL;
    bipolar        : BOOL;
    measuringMode  : INT;
    retVal         : WORD;
    outputValue    : REAL;
END_STRUCT
END_TYPE;

FUNCTION_BLOCK FB_AnalogBatchProcessing
VAR_INPUT
    count : DINT;
END_VAR
VAR_IN_OUT
    analogValues : ARRAY[*] OF INT;
    channels     : ARRAY[*] OF ST_AnalogChannel;
END_VAR
VAR_OUTPUT
END_VAR
VAR
END_VAR

(*
ENGINEERING_CONTRACT
================================================================================
PUB001: Process 'count' channels starting at each array's lower bound.
        Arrays passed by reference preserve caller-defined bounds.
        Read-only: analogValues elements are never modified.
PUB002: Per-channel conversion based on measuringMode field.
        - Mode 0: Linear scaling using hiLIM/loLIM and bipolar flag.
        - Mode 1: Standard temperature (raw / 10.0).
        - Mode 2: Climatic temperature (raw / 100.0).
        - Invalid mode: retVal=16#8001, outputValue unchanged.
PUB003: Mode 0 linear scaling maps raw 0..27648 (unipolar) or -27648..27648 (bipolar)
        to loLIM..hiLIM range. OutputValue = loLIM + (raw - rawMin) * (hiLIM - loLIM) / range.
PUB004: If hiLIM <= loLIM in mode 0, set retVal=16#8002 and skip conversion.
PUB005: Disabled channels (enable=FALSE) are skipped; retVal and outputValue unchanged.
PUB006: Per-channel retVal WORD status: 16#8001 (invalid mode), 16#8002 (bad range).
PUB007: Same-scan priority: enable→measuringMode→hiLIM/loLIM check→conversion.
PUB008: Temperature output = raw / divisor (10 or 100) as REAL.
--------------------------------------------------------------------------------
*)

VAR
    tmpIndex     : DINT;
    tmpRaw       : INT;
    tmpRawReal   : REAL;
    tmpRange     : REAL;
    tmpOffset    : REAL;
    tmpChannel   : ST_AnalogChannel;
    tmpLower     : DINT;
    tmpUpperAna  : DINT;
    tmpUpperCh   : DINT;
    tmpProcessed : BOOL;
END_VAR

(* CONTRACT_RULES [] *)

tmpLower    := LOWER_BOUND(analogValues, 1);
tmpUpperAna := UPPER_BOUND(analogValues, 1);
tmpUpperCh  := UPPER_BOUND(channels, 1);

FOR tmpIndex := 0 TO (count - 1) DO
    tmpProcessed := FALSE;

    (* Bounds check: skip if index exceeds either array *)
    IF (tmpLower + tmpIndex) <= tmpUpperAna AND (tmpLower + tmpIndex) <= tmpUpperCh THEN
        tmpChannel := channels[tmpLower + tmpIndex];

        (* Skip disabled channels; retain previous outputValue and retVal *)
        IF tmpChannel.enable THEN

    (* Determine conversion based on measuringMode *)
    IF tmpChannel.measuringMode = 0 THEN
        (* Non-temperature linear scaling *)
        IF tmpChannel.hiLIM <= tmpChannel.loLIM THEN
            channels[tmpLower + tmpIndex].retVal := 16#8002;
        ELSE
            tmpRaw       := analogValues[tmpLower + tmpIndex];
            tmpRawReal   := TO_REAL(tmpRaw);
            tmpRange     := tmpChannel.hiLIM - tmpChannel.loLIM;

            IF tmpChannel.bipolar THEN
                (* Map -27648..27648 to loLIM..hiLIM *)
                tmpOffset    := TO_REAL(27648);
                channels[tmpLower + tmpIndex].outputValue := tmpChannel.loLIM +
                    (tmpRawReal + tmpOffset) * tmpRange / TO_REAL(55296);
            ELSE
                (* Map 0..27648 to loLIM..hiLIM *)
                channels[tmpLower + tmpIndex].outputValue := tmpChannel.loLIM +
                    tmpRawReal * tmpRange / TO_REAL(27648);
            END_IF;
            channels[tmpLower + tmpIndex].retVal := 0;
        END_IF;
        tmpProcessed := TRUE;
    ELSIF tmpChannel.measuringMode = 1 THEN
        (* Standard temperature: outputValue = raw / 10 *)
        tmpRaw := analogValues[tmpLower + tmpIndex];
        channels[tmpLower + tmpIndex].outputValue := TO_REAL(tmpRaw) / TO_REAL(10);
        channels[tmpLower + tmpIndex].retVal := 0;
        tmpProcessed := TRUE;
    ELSIF tmpChannel.measuringMode = 2 THEN
        (* Climatic temperature: outputValue = raw / 100 *)
        tmpRaw := analogValues[tmpLower + tmpIndex];
        channels[tmpLower + tmpIndex].outputValue := TO_REAL(tmpRaw) / TO_REAL(100);
        channels[tmpLower + tmpIndex].retVal := 0;
        tmpProcessed := TRUE;
    END_IF;

    (* Invalid measuringMode (not 0, 1, or 2) *)
    IF NOT tmpProcessed THEN
        channels[tmpLower + tmpIndex].retVal := 16#8001;
    END_IF;

END_FOR;

END_FUNCTION_BLOCK

(* ---- public-medium-02.candidate_03.st ---- *)
TYPE ST_AnalogChannel :
STRUCT
    enable         : BOOL;
    hiLIM          : REAL;
    loLIM          : REAL;
    bipolar        : BOOL;
    measuringMode  : INT;
    retVal         : WORD;
    outputValue    : REAL;
END_STRUCT
END_TYPE;

FUNCTION_BLOCK FB_AnalogBatchProcessing
VAR_INPUT
    count : DINT;
END_VAR
VAR_IN_OUT
    analogValues : ARRAY[*] OF INT;
    channels     : ARRAY[*] OF ST_AnalogChannel;
END_VAR
VAR_OUTPUT
END_VAR
VAR
END_VAR

(*
ENGINEERING_CONTRACT
================================================================================
PUB001: Process 'count' channels starting at each array's lower bound.
        Arrays passed by reference preserve caller-defined bounds.
        Read-only: analogValues elements are never modified.
PUB002: Per-channel conversion based on measuringMode field.
        - Mode 0: Linear scaling using hiLIM/loLIM and bipolar flag.
        - Mode 1: Standard temperature (raw / 10.0).
        - Mode 2: Climatic temperature (raw / 100.0).
        - Invalid mode: retVal=16#8001, outputValue unchanged.
PUB003: Mode 0 linear scaling maps raw 0..27648 (unipolar) or -27648..27648 (bipolar)
        to loLIM..hiLIM range. OutputValue = loLIM + (raw - rawMin) * (hiLIM - loLIM) / range.
PUB004: If hiLIM <= loLIM in mode 0, set retVal=16#8002 and skip conversion.
PUB005: Disabled channels (enable=FALSE) are skipped; retVal and outputValue unchanged.
PUB006: Per-channel retVal WORD status: 16#8001 (invalid mode), 16#8002 (bad range).
PUB007: Same-scan priority: enable→measuringMode→hiLIM/loLIM check→conversion.
PUB008: Temperature output = raw / divisor (10 or 100) as REAL.
--------------------------------------------------------------------------------
*)

VAR
    tmpIndex     : DINT;
    tmpRaw       : INT;
    tmpRawReal   : REAL;
    tmpRange     : REAL;
    tmpOffset    : REAL;
    tmpChannel   : ST_AnalogChannel;
    tmpLower     : DINT;
    tmpUpperAna  : DINT;
    tmpUpperCh   : DINT;
    tmpProcessed : BOOL;
END_VAR

(* CONTRACT_RULES [] *)

tmpLower    := LOWER_BOUND(analogValues, 1);
tmpUpperAna := UPPER_BOUND(analogValues, 1);
tmpUpperCh  := UPPER_BOUND(channels, 1);

FOR tmpIndex := 0 TO (count - 1) DO
    tmpProcessed := FALSE;

    (* Bounds check: skip if index exceeds either array *)
    IF (tmpLower + tmpIndex) <= tmpUpperAna AND (tmpLower + tmpIndex) <= tmpUpperCh THEN
        tmpChannel := channels[tmpLower + tmpIndex];

        (* Skip disabled channels; retain previous outputValue and retVal *)
        IF tmpChannel.enable THEN

    (* Determine conversion based on measuringMode *)
    IF tmpChannel.measuringMode = 0 THEN
        (* Non-temperature linear scaling *)
        IF tmpChannel.hiLIM <= tmpChannel.loLIM THEN
            channels[tmpLower + tmpIndex].retVal := 16#8002;
        ELSE
            tmpRaw       := analogValues[tmpLower + tmpIndex];
            tmpRawReal   := TO_REAL(tmpRaw);
            tmpRange     := tmpChannel.hiLIM - tmpChannel.loLIM;

            IF tmpChannel.bipolar THEN
                (* Map -27648..27648 to loLIM..hiLIM *)
                tmpOffset    := TO_REAL(27648);
                channels[tmpLower + tmpIndex].outputValue := tmpChannel.loLIM +
                    (tmpRawReal + tmpOffset) * tmpRange / TO_REAL(55296);
            ELSE
                (* Map 0..27648 to loLIM..hiLIM *)
                channels[tmpLower + tmpIndex].outputValue := tmpChannel.loLIM +
                    tmpRawReal * tmpRange / TO_REAL(27648);
            END_IF;
            channels[tmpLower + tmpIndex].retVal := 0;
        END_IF;
        tmpProcessed := TRUE;
    ELSIF tmpChannel.measuringMode = 1 THEN
        (* Standard temperature: outputValue = raw / 10 *)
        tmpRaw := analogValues[tmpLower + tmpIndex];
        channels[tmpLower + tmpIndex].outputValue := TO_REAL(tmpRaw) / TO_REAL(10);
        channels[tmpLower + tmpIndex].retVal := 0;
        tmpProcessed := TRUE;
    ELSIF tmpChannel.measuringMode = 2 THEN
        (* Climatic temperature: outputValue = raw / 100 *)
        tmpRaw := analogValues[tmpLower + tmpIndex];
        channels[tmpLower + tmpIndex].outputValue := TO_REAL(tmpRaw) / TO_REAL(100);
        channels[tmpLower + tmpIndex].retVal := 0;
        tmpProcessed := TRUE;
    END_IF;

    (* Invalid measuringMode (not 0, 1, or 2) *)
    IF NOT tmpProcessed THEN
        channels[tmpLower + tmpIndex].retVal := 16#8001;
    END_IF;

    END_IF; (* close outer enable check *)

END_FOR;

END_FUNCTION_BLOCK

(* ---- public-medium-02.patch_base_02.st ---- *)
FUNCTION_BLOCK FB_AnalogBatchProcessing
VAR_INPUT
END_VAR
VAR_IN_OUT
    analogValues : ARRAY[*] OF INT;
    channels     : ARRAY[*] OF ST_AnalogChannel;
END_VAR
VAR_OUTPUT
END_VAR
VAR
END_VAR

(*
ENGINEERING_CONTRACT
================================================================================
PUB001: Process 'count' channels starting at each array's lower bound.
        Arrays passed by reference preserve caller-defined bounds.
        Read-only: analogValues elements are never modified.
PUB002: Per-channel conversion based on measuringMode field.
        - Mode 0: Linear scaling using hiLIM/loLIM and bipolar flag.
        - Mode 1: Standard temperature (raw / 10.0).
        - Mode 2: Climatic temperature (raw / 100.0).
        - Invalid mode: retVal=16#8001, outputValue unchanged.
PUB003: Mode 0 linear scaling maps raw 0..27648 (unipolar) or -27648..27648 (bipolar)
        to loLIM..hiLIM range. OutputValue = loLIM + (raw - rawMin) * (hiLIM - loLIM) / range.
PUB004: If hiLIM <= loLIM in mode 0, set retVal=16#8002 and skip conversion.
PUB005: Disabled channels (enable=FALSE) are skipped; retVal and outputValue unchanged.
PUB006: Per-channel retVal WORD status: 16#8001 (invalid mode), 16#8002 (bad range).
PUB007: Same-scan priority: enable→measuringMode→hiLIM/loLIM check→conversion.
PUB008: Temperature output = raw / divisor (10 or 100) as REAL.
--------------------------------------------------------------------------------
*)

VAR
    tmpIndex     : DINT;
    tmpRaw       : INT;
    tmpRawReal   : REAL;
    tmpRange     : REAL;
    tmpOffset    : REAL;
    tmpChannel   : ST_AnalogChannel;
    tmpLower     : DINT;
    tmpUpperAna  : DINT;
    tmpUpperCh   : DINT;
    tmpProcessed : BOOL;
END_VAR

(* CONTRACT_RULES [] *)

tmpLower    := LOWER_BOUND(analogValues, 1);
tmpUpperAna := UPPER_BOUND(analogValues, 1);
tmpUpperCh  := UPPER_BOUND(channels, 1);

FOR tmpIndex := 0 TO (count - 1) DO
    tmpProcessed := FALSE;

    (* Bounds check: skip if index exceeds either array *)
    IF (tmpLower + tmpIndex) > tmpUpperAna OR (tmpLower + tmpIndex) > tmpUpperCh THEN
        CONTINUE;
    END_IF;

    tmpChannel := channels[tmpLower + tmpIndex];

    (* Skip disabled channels; retain previous outputValue and retVal *)
    IF NOT tmpChannel.enable THEN
        CONTINUE;
    END_IF;

    (* Determine conversion based on measuringMode *)
    IF tmpChannel.measuringMode = 0 THEN
        (* Non-temperature linear scaling *)
        IF tmpChannel.hiLIM <= tmpChannel.loLIM THEN
            channels[tmpLower + tmpIndex].retVal := 16#8002;
        ELSE
            tmpRaw       := analogValues[tmpLower + tmpIndex];
            tmpRawReal   := TO_REAL(tmpRaw);
            tmpRange     := tmpChannel.hiLIM - tmpChannel.loLIM;

            IF tmpChannel.bipolar THEN
                (* Map -27648..27648 to loLIM..hiLIM *)
                tmpOffset    := TO_REAL(27648);
                channels[tmpLower + tmpIndex].outputValue := tmpChannel.loLIM +
                    (tmpRawReal + tmpOffset) * tmpRange / TO_REAL(55296);
            ELSE
                (* Map 0..27648 to loLIM..hiLIM *)
                channels[tmpLower + tmpIndex].outputValue := tmpChannel.loLIM +
                    tmpRawReal * tmpRange / TO_REAL(27648);
            END_IF;
            channels[tmpLower + tmpIndex].retVal := 0;
        END_IF;
        tmpProcessed := TRUE;
    ELSIF tmpChannel.measuringMode = 1 THEN
        (* Standard temperature: outputValue = raw / 10 *)
        tmpRaw := analogValues[tmpLower + tmpIndex];
        channels[tmpLower + tmpIndex].outputValue := TO_REAL(tmpRaw) / TO_REAL(10);
        channels[tmpLower + tmpIndex].retVal := 0;
        tmpProcessed := TRUE;
    ELSIF tmpChannel.measuringMode = 2 THEN
        (* Climatic temperature: outputValue = raw / 100 *)
        tmpRaw := analogValues[tmpLower + tmpIndex];
        channels[tmpLower + tmpIndex].outputValue := TO_REAL(tmpRaw) / TO_REAL(100);
        channels[tmpLower + tmpIndex].retVal := 0;
        tmpProcessed := TRUE;
    END_IF;

    (* Invalid measuringMode (not 0, 1, or 2) *)
    IF NOT tmpProcessed THEN
        channels[tmpLower + tmpIndex].retVal := 16#8001;
    END_IF;

END_FOR;

END_FUNCTION_BLOCK

(* ---- public-medium-02.patch_base_03.st ---- *)
TYPE ST_AnalogChannel :
STRUCT
    enable         : BOOL;
    hiLIM          : REAL;
    loLIM          : REAL;
    bipolar        : BOOL;
    measuringMode  : INT;
    retVal         : WORD;
    outputValue    : REAL;
END_STRUCT
END_TYPE;

FUNCTION_BLOCK FB_AnalogBatchProcessing
VAR_INPUT
    count : DINT;
END_VAR
VAR_IN_OUT
    analogValues : ARRAY[*] OF INT;
    channels     : ARRAY[*] OF ST_AnalogChannel;
END_VAR
VAR_OUTPUT
END_VAR
VAR
END_VAR

(*
ENGINEERING_CONTRACT
================================================================================
PUB001: Process 'count' channels starting at each array's lower bound.
        Arrays passed by reference preserve caller-defined bounds.
        Read-only: analogValues elements are never modified.
PUB002: Per-channel conversion based on measuringMode field.
        - Mode 0: Linear scaling using hiLIM/loLIM and bipolar flag.
        - Mode 1: Standard temperature (raw / 10.0).
        - Mode 2: Climatic temperature (raw / 100.0).
        - Invalid mode: retVal=16#8001, outputValue unchanged.
PUB003: Mode 0 linear scaling maps raw 0..27648 (unipolar) or -27648..27648 (bipolar)
        to loLIM..hiLIM range. OutputValue = loLIM + (raw - rawMin) * (hiLIM - loLIM) / range.
PUB004: If hiLIM <= loLIM in mode 0, set retVal=16#8002 and skip conversion.
PUB005: Disabled channels (enable=FALSE) are skipped; retVal and outputValue unchanged.
PUB006: Per-channel retVal WORD status: 16#8001 (invalid mode), 16#8002 (bad range).
PUB007: Same-scan priority: enable→measuringMode→hiLIM/loLIM check→conversion.
PUB008: Temperature output = raw / divisor (10 or 100) as REAL.
--------------------------------------------------------------------------------
*)

VAR
    tmpIndex     : DINT;
    tmpRaw       : INT;
    tmpRawReal   : REAL;
    tmpRange     : REAL;
    tmpOffset    : REAL;
    tmpChannel   : ST_AnalogChannel;
    tmpLower     : DINT;
    tmpUpperAna  : DINT;
    tmpUpperCh   : DINT;
    tmpProcessed : BOOL;
END_VAR

(* CONTRACT_RULES [] *)

tmpLower    := LOWER_BOUND(analogValues, 1);
tmpUpperAna := UPPER_BOUND(analogValues, 1);
tmpUpperCh  := UPPER_BOUND(channels, 1);

FOR tmpIndex := 0 TO (count - 1) DO
    tmpProcessed := FALSE;

    (* Bounds check: skip if index exceeds either array *)
    IF (tmpLower + tmpIndex) <= tmpUpperAna AND (tmpLower + tmpIndex) <= tmpUpperCh THEN
        tmpChannel := channels[tmpLower + tmpIndex];

        (* Skip disabled channels; retain previous outputValue and retVal *)
        IF tmpChannel.enable THEN

    (* Determine conversion based on measuringMode *)
    IF tmpChannel.measuringMode = 0 THEN
        (* Non-temperature linear scaling *)
        IF tmpChannel.hiLIM <= tmpChannel.loLIM THEN
            channels[tmpLower + tmpIndex].retVal := 16#8002;
        ELSE
            tmpRaw       := analogValues[tmpLower + tmpIndex];
            tmpRawReal   := TO_REAL(tmpRaw);
            tmpRange     := tmpChannel.hiLIM - tmpChannel.loLIM;

            IF tmpChannel.bipolar THEN
                (* Map -27648..27648 to loLIM..hiLIM *)
                tmpOffset    := TO_REAL(27648);
                channels[tmpLower + tmpIndex].outputValue := tmpChannel.loLIM +
                    (tmpRawReal + tmpOffset) * tmpRange / TO_REAL(55296);
            ELSE
                (* Map 0..27648 to loLIM..hiLIM *)
                channels[tmpLower + tmpIndex].outputValue := tmpChannel.loLIM +
                    tmpRawReal * tmpRange / TO_REAL(27648);
            END_IF;
            channels[tmpLower + tmpIndex].retVal := 0;
        END_IF;
        tmpProcessed := TRUE;
    ELSIF tmpChannel.measuringMode = 1 THEN
        (* Standard temperature: outputValue = raw / 10 *)
        tmpRaw := analogValues[tmpLower + tmpIndex];
        channels[tmpLower + tmpIndex].outputValue := TO_REAL(tmpRaw) / TO_REAL(10);
        channels[tmpLower + tmpIndex].retVal := 0;
        tmpProcessed := TRUE;
    ELSIF tmpChannel.measuringMode = 2 THEN
        (* Climatic temperature: outputValue = raw / 100 *)
        tmpRaw := analogValues[tmpLower + tmpIndex];
        channels[tmpLower + tmpIndex].outputValue := TO_REAL(tmpRaw) / TO_REAL(100);
        channels[tmpLower + tmpIndex].retVal := 0;
        tmpProcessed := TRUE;
    END_IF;

    (* Invalid measuringMode (not 0, 1, or 2) *)
    IF NOT tmpProcessed THEN
        channels[tmpLower + tmpIndex].retVal := 16#8001;
    END_IF;

END_FOR;

END_FUNCTION_BLOCK

(* ---- public-medium-02.patch_base_04.st ---- *)
TYPE ST_AnalogChannel :
STRUCT
    enable         : BOOL;
    hiLIM          : REAL;
    loLIM          : REAL;
    bipolar        : BOOL;
    measuringMode  : INT;
    retVal         : WORD;
    outputValue    : REAL;
END_STRUCT
END_TYPE;

FUNCTION_BLOCK FB_AnalogBatchProcessing
VAR_INPUT
    count : DINT;
END_VAR
VAR_IN_OUT
    analogValues : ARRAY[*] OF INT;
    channels     : ARRAY[*] OF ST_AnalogChannel;
END_VAR
VAR_OUTPUT
END_VAR
VAR
END_VAR

(*
ENGINEERING_CONTRACT
================================================================================
PUB001: Process 'count' channels starting at each array's lower bound.
        Arrays passed by reference preserve caller-defined bounds.
        Read-only: analogValues elements are never modified.
PUB002: Per-channel conversion based on measuringMode field.
        - Mode 0: Linear scaling using hiLIM/loLIM and bipolar flag.
        - Mode 1: Standard temperature (raw / 10.0).
        - Mode 2: Climatic temperature (raw / 100.0).
        - Invalid mode: retVal=16#8001, outputValue unchanged.
PUB003: Mode 0 linear scaling maps raw 0..27648 (unipolar) or -27648..27648 (bipolar)
        to loLIM..hiLIM range. OutputValue = loLIM + (raw - rawMin) * (hiLIM - loLIM) / range.
PUB004: If hiLIM <= loLIM in mode 0, set retVal=16#8002 and skip conversion.
PUB005: Disabled channels (enable=FALSE) are skipped; retVal and outputValue unchanged.
PUB006: Per-channel retVal WORD status: 16#8001 (invalid mode), 16#8002 (bad range).
PUB007: Same-scan priority: enable→measuringMode→hiLIM/loLIM check→conversion.
PUB008: Temperature output = raw / divisor (10 or 100) as REAL.
--------------------------------------------------------------------------------
*)

VAR
    tmpIndex     : DINT;
    tmpRaw       : INT;
    tmpRawReal   : REAL;
    tmpRange     : REAL;
    tmpOffset    : REAL;
    tmpChannel   : ST_AnalogChannel;
    tmpLower     : DINT;
    tmpUpperAna  : DINT;
    tmpUpperCh   : DINT;
    tmpProcessed : BOOL;
END_VAR

(* CONTRACT_RULES [] *)

tmpLower    := LOWER_BOUND(analogValues, 1);
tmpUpperAna := UPPER_BOUND(analogValues, 1);
tmpUpperCh  := UPPER_BOUND(channels, 1);

FOR tmpIndex := 0 TO (count - 1) DO
    tmpProcessed := FALSE;

    (* Bounds check: skip if index exceeds either array *)
    IF (tmpLower + tmpIndex) <= tmpUpperAna AND (tmpLower + tmpIndex) <= tmpUpperCh THEN
        tmpChannel := channels[tmpLower + tmpIndex];

        (* Skip disabled channels; retain previous outputValue and retVal *)
        IF tmpChannel.enable THEN

    (* Determine conversion based on measuringMode *)
    IF tmpChannel.measuringMode = 0 THEN
        (* Non-temperature linear scaling *)
        IF tmpChannel.hiLIM <= tmpChannel.loLIM THEN
            channels[tmpLower + tmpIndex].retVal := 16#8002;
        ELSE
            tmpRaw       := analogValues[tmpLower + tmpIndex];
            tmpRawReal   := TO_REAL(tmpRaw);
            tmpRange     := tmpChannel.hiLIM - tmpChannel.loLIM;

            IF tmpChannel.bipolar THEN
                (* Map -27648..27648 to loLIM..hiLIM *)
                tmpOffset    := TO_REAL(27648);
                channels[tmpLower + tmpIndex].outputValue := tmpChannel.loLIM +
                    (tmpRawReal + tmpOffset) * tmpRange / TO_REAL(55296);
            ELSE
                (* Map 0..27648 to loLIM..hiLIM *)
                channels[tmpLower + tmpIndex].outputValue := tmpChannel.loLIM +
                    tmpRawReal * tmpRange / TO_REAL(27648);
            END_IF;
            channels[tmpLower + tmpIndex].retVal := 0;
        END_IF;
        tmpProcessed := TRUE;
    ELSIF tmpChannel.measuringMode = 1 THEN
        (* Standard temperature: outputValue = raw / 10 *)
        tmpRaw := analogValues[tmpLower + tmpIndex];
        channels[tmpLower + tmpIndex].outputValue := TO_REAL(tmpRaw) / TO_REAL(10);
        channels[tmpLower + tmpIndex].retVal := 0;
        tmpProcessed := TRUE;
    ELSIF tmpChannel.measuringMode = 2 THEN
        (* Climatic temperature: outputValue = raw / 100 *)
        tmpRaw := analogValues[tmpLower + tmpIndex];
        channels[tmpLower + tmpIndex].outputValue := TO_REAL(tmpRaw) / TO_REAL(100);
        channels[tmpLower + tmpIndex].retVal := 0;
        tmpProcessed := TRUE;
    END_IF;

    (* Invalid measuringMode (not 0, 1, or 2) *)
    IF NOT tmpProcessed THEN
        channels[tmpLower + tmpIndex].retVal := 16#8001;
    END_IF;

    END_IF; (* close outer enable check *)

END_FOR;

END_FUNCTION_BLOCK

(* ---- public-medium-02.raw_candidate_01.st ---- *)
FUNCTION_BLOCK FB_AnalogBatchProcessing
VAR_INPUT
END_VAR
VAR_IN_OUT
    analogValues : ARRAY[*] OF INT;
    channels     : ARRAY[*] OF ST_AnalogChannel;
END_VAR
VAR_OUTPUT
END_VAR
VAR
END_VAR

(*
ENGINEERING_CONTRACT
================================================================================
PUB001: Process 'count' channels starting at each array's lower bound.
        Arrays passed by reference preserve caller-defined bounds.
        Read-only: analogValues elements are never modified.
PUB002: Per-channel conversion based on measuringMode field.
        - Mode 0: Linear scaling using hiLIM/loLIM and bipolar flag.
        - Mode 1: Standard temperature (raw / 10.0).
        - Mode 2: Climatic temperature (raw / 100.0).
        - Invalid mode: retVal=16#8001, outputValue unchanged.
PUB003: Mode 0 linear scaling maps raw 0..27648 (unipolar) or -27648..27648 (bipolar)
        to loLIM..hiLIM range. OutputValue = loLIM + (raw - rawMin) * (hiLIM - loLIM) / range.
PUB004: If hiLIM <= loLIM in mode 0, set retVal=16#8002 and skip conversion.
PUB005: Disabled channels (enable=FALSE) are skipped; retVal and outputValue unchanged.
PUB006: Per-channel retVal WORD status: 16#8001 (invalid mode), 16#8002 (bad range).
PUB007: Same-scan priority: enable→measuringMode→hiLIM/loLIM check→conversion.
PUB008: Temperature output = raw / divisor (10 or 100) as REAL.
--------------------------------------------------------------------------------
*)

VAR
    tmpIndex     : DINT;
    tmpRaw       : INT;
    tmpRawReal   : REAL;
    tmpRange     : REAL;
    tmpOffset    : REAL;
    tmpChannel   : ST_AnalogChannel;
    tmpLower     : DINT;
    tmpUpperAna  : DINT;
    tmpUpperCh   : DINT;
    tmpProcessed : BOOL;
END_VAR

(* CONTRACT_RULES [] *)

tmpLower    := LOWER_BOUND(analogValues, 1);
tmpUpperAna := UPPER_BOUND(analogValues, 1);
tmpUpperCh  := UPPER_BOUND(channels, 1);

FOR tmpIndex := 0 TO (count - 1) DO
    tmpProcessed := FALSE;

    (* Bounds check: skip if index exceeds either array *)
    IF (tmpLower + tmpIndex) > tmpUpperAna OR (tmpLower + tmpIndex) > tmpUpperCh THEN
        CONTINUE;
    END_IF

    tmpChannel := channels[tmpLower + tmpIndex];

    (* Skip disabled channels; retain previous outputValue and retVal *)
    IF NOT tmpChannel.enable THEN
        CONTINUE;
    END_IF

    (* Determine conversion based on measuringMode *)
    IF tmpChannel.measuringMode = 0 THEN
        (* Non-temperature linear scaling *)
        IF tmpChannel.hiLIM <= tmpChannel.loLIM THEN
            channels[tmpLower + tmpIndex].retVal := 16#8002;
        ELSE
            tmpRaw       := analogValues[tmpLower + tmpIndex];
            tmpRawReal   := TO_REAL(tmpRaw);
            tmpRange     := tmpChannel.hiLIM - tmpChannel.loLIM;

            IF tmpChannel.bipolar THEN
                (* Map -27648..27648 to loLIM..hiLIM *)
                tmpOffset    := TO_REAL(27648);
                channels[tmpLower + tmpIndex].outputValue := tmpChannel.loLIM +
                    (tmpRawReal + tmpOffset) * tmpRange / TO_REAL(55296);
            ELSE
                (* Map 0..27648 to loLIM..hiLIM *)
                channels[tmpLower + tmpIndex].outputValue := tmpChannel.loLIM +
                    tmpRawReal * tmpRange / TO_REAL(27648);
            END_IF
            channels[tmpLower + tmpIndex].retVal := 0;
        END_IF
        tmpProcessed := TRUE;
    ELSIF tmpChannel.measuringMode = 1 THEN
        (* Standard temperature: outputValue = raw / 10 *)
        tmpRaw := analogValues[tmpLower + tmpIndex];
        channels[tmpLower + tmpIndex].outputValue := TO_REAL(tmpRaw) / TO_REAL(10);
        channels[tmpLower + tmpIndex].retVal := 0;
        tmpProcessed := TRUE;
    ELSIF tmpChannel.measuringMode = 2 THEN
        (* Climatic temperature: outputValue = raw / 100 *)
        tmpRaw := analogValues[tmpLower + tmpIndex];
        channels[tmpLower + tmpIndex].outputValue := TO_REAL(tmpRaw) / TO_REAL(100);
        channels[tmpLower + tmpIndex].retVal := 0;
        tmpProcessed := TRUE;
    END_IF

    (* Invalid measuringMode (not 0, 1, or 2) *)
    IF NOT tmpProcessed THEN
        channels[tmpLower + tmpIndex].retVal := 16#8001;
    END_IF

END_FOR;

END_FUNCTION_BLOCK

(* ---- public-medium-02.raw_candidate_02.st ---- *)
TYPE ST_AnalogChannel :
STRUCT
    enable         : BOOL;
    hiLIM          : REAL;
    loLIM          : REAL;
    bipolar        : BOOL;
    measuringMode  : INT;
    retVal         : WORD;
    outputValue    : REAL;
END_STRUCT
END_TYPE

FUNCTION_BLOCK FB_AnalogBatchProcessing
VAR_INPUT
    count : DINT;
END_VAR
VAR_IN_OUT
    analogValues : ARRAY[*] OF INT;
    channels     : ARRAY[*] OF ST_AnalogChannel;
END_VAR
VAR_OUTPUT
END_VAR
VAR
END_VAR

(*
ENGINEERING_CONTRACT
================================================================================
PUB001: Process 'count' channels starting at each array's lower bound.
        Arrays passed by reference preserve caller-defined bounds.
        Read-only: analogValues elements are never modified.
PUB002: Per-channel conversion based on measuringMode field.
        - Mode 0: Linear scaling using hiLIM/loLIM and bipolar flag.
        - Mode 1: Standard temperature (raw / 10.0).
        - Mode 2: Climatic temperature (raw / 100.0).
        - Invalid mode: retVal=16#8001, outputValue unchanged.
PUB003: Mode 0 linear scaling maps raw 0..27648 (unipolar) or -27648..27648 (bipolar)
        to loLIM..hiLIM range. OutputValue = loLIM + (raw - rawMin) * (hiLIM - loLIM) / range.
PUB004: If hiLIM <= loLIM in mode 0, set retVal=16#8002 and skip conversion.
PUB005: Disabled channels (enable=FALSE) are skipped; retVal and outputValue unchanged.
PUB006: Per-channel retVal WORD status: 16#8001 (invalid mode), 16#8002 (bad range).
PUB007: Same-scan priority: enable→measuringMode→hiLIM/loLIM check→conversion.
PUB008: Temperature output = raw / divisor (10 or 100) as REAL.
--------------------------------------------------------------------------------
*)

VAR
    tmpIndex     : DINT;
    tmpRaw       : INT;
    tmpRawReal   : REAL;
    tmpRange     : REAL;
    tmpOffset    : REAL;
    tmpChannel   : ST_AnalogChannel;
    tmpLower     : DINT;
    tmpUpperAna  : DINT;
    tmpUpperCh   : DINT;
    tmpProcessed : BOOL;
END_VAR

(* CONTRACT_RULES [] *)

tmpLower    := LOWER_BOUND(analogValues, 1);
tmpUpperAna := UPPER_BOUND(analogValues, 1);
tmpUpperCh  := UPPER_BOUND(channels, 1);

FOR tmpIndex := 0 TO (count - 1) DO
    tmpProcessed := FALSE;

    (* Bounds check: skip if index exceeds either array *)
    IF (tmpLower + tmpIndex) <= tmpUpperAna AND (tmpLower + tmpIndex) <= tmpUpperCh THEN
        tmpChannel := channels[tmpLower + tmpIndex];

        (* Skip disabled channels; retain previous outputValue and retVal *)
        IF tmpChannel.enable THEN

    (* Determine conversion based on measuringMode *)
    IF tmpChannel.measuringMode = 0 THEN
        (* Non-temperature linear scaling *)
        IF tmpChannel.hiLIM <= tmpChannel.loLIM THEN
            channels[tmpLower + tmpIndex].retVal := 16#8002;
        ELSE
            tmpRaw       := analogValues[tmpLower + tmpIndex];
            tmpRawReal   := TO_REAL(tmpRaw);
            tmpRange     := tmpChannel.hiLIM - tmpChannel.loLIM;

            IF tmpChannel.bipolar THEN
                (* Map -27648..27648 to loLIM..hiLIM *)
                tmpOffset    := TO_REAL(27648);
                channels[tmpLower + tmpIndex].outputValue := tmpChannel.loLIM +
                    (tmpRawReal + tmpOffset) * tmpRange / TO_REAL(55296);
            ELSE
                (* Map 0..27648 to loLIM..hiLIM *)
                channels[tmpLower + tmpIndex].outputValue := tmpChannel.loLIM +
                    tmpRawReal * tmpRange / TO_REAL(27648);
            END_IF;
            channels[tmpLower + tmpIndex].retVal := 0;
        END_IF;
        tmpProcessed := TRUE;
    ELSIF tmpChannel.measuringMode = 1 THEN
        (* Standard temperature: outputValue = raw / 10 *)
        tmpRaw := analogValues[tmpLower + tmpIndex];
        channels[tmpLower + tmpIndex].outputValue := TO_REAL(tmpRaw) / TO_REAL(10);
        channels[tmpLower + tmpIndex].retVal := 0;
        tmpProcessed := TRUE;
    ELSIF tmpChannel.measuringMode = 2 THEN
        (* Climatic temperature: outputValue = raw / 100 *)
        tmpRaw := analogValues[tmpLower + tmpIndex];
        channels[tmpLower + tmpIndex].outputValue := TO_REAL(tmpRaw) / TO_REAL(100);
        channels[tmpLower + tmpIndex].retVal := 0;
        tmpProcessed := TRUE;
    END_IF;

    (* Invalid measuringMode (not 0, 1, or 2) *)
    IF NOT tmpProcessed THEN
        channels[tmpLower + tmpIndex].retVal := 16#8001;
    END_IF;

END_FOR;

END_FUNCTION_BLOCK
